def _start_heartbeat():
    import threading as _t, time as _time, os as _os, io as _io
    def _beat():
        while True:
            try:
                last = ''
                try:
                    with _io.open(LOG_PATH, 'r', encoding='utf-8') as f:
                        _lines = f.read().splitlines()
                        last = _lines[-1] if _lines else ''
                except Exception:
                    pass
                with _io.open(HEARTBEAT_PATH, 'w', encoding='utf-8') as f:
                    f.write('%s | pid=%d | alive\nlast: %s\n' % (
                        _time.strftime('%m-%d %H:%M:%S'), _os.getpid(), last[:150]))
            except Exception:
                pass
            _time.sleep(5.0)
    _t.Thread(target=_beat, daemon=True, name='gui_heartbeat').start()


def log(s):
    _file_log(s)  # 先落盘：即使后续 print 阻塞，磁盘日志也不受影响
    print(s)
    if text_log:
        try:
            _log_queue.put_nowait(str(s))
        except Exception:
            text_log.insert(tk.END, str(s) + NL)

# ============================================================
# 连接（只连一次，复用）
# ============================================================
def ensure_connected():
    global _connected
    try:
        status, msg = robot.ConnectedState()
        if status != ROBOTCOM_READY:
            if status >= 0:
                log('机器人未就绪，取消执行：' + str(msg))
                return False
            robot.Connect()
            # v14o：固定 1.5s 改为就绪探测（0.3s 轮询，最多 3s）：假断连恢复是每跳尾部
            # 停顿税的一部分；探测到就绪即返回，未就绪语义与旧版一致（返回 False）。
            for _ in range(10):
                time.sleep(0.3)
                status, msg = robot.ConnectedState()
                if status == ROBOTCOM_READY:
                    break
        _connected = status == ROBOTCOM_READY
        if not _connected:
            log('机器人连接未就绪：' + str(msg))
            return False
        RDK.setRunMode(RUNMODE_RUN_ROBOT)
        return True
    except Exception as exc:
        _connected = False
        log('连接失败：' + str(exc))
        return False


# ============================================================
# 解析坐标
# ============================================================
def parse_points():
    if not text_points:
        return []
    raw = text_points.get("1.0", tk.END)
    points = []
    for line in raw.strip().split(NL):
        line = line.strip()
        if not line or line.startswith("#"):
            continue
        try:
            vals = [float(v.strip()) for v in line.split(",")]
            if len(vals) >= 6:
                points.append(vals[:6])
        except ValueError:
            pass
    return points

# ============================================================
# 读取当前位置
# ============================================================
def read_current(entries=None):
    try:
        pose = robot.Pose()
        v = pose_to_fanuc(pose)
        log("")
        log("当前 TCP：X=%.3f Y=%.3f Z=%.3f Rx=%.3f Ry=%.3f Rz=%.3f" % tuple(v[:6]))
    except Exception as e:
        log("读取失败：%s" % e)

def fill_current(entries=None):
    try:
        pose = robot.Pose()
        v = pose_to_fanuc(pose)
        if entries:
            for e, val in zip(entries, v):
                e.delete(0, tk.END)
                e.insert(0, "%.3f" % val)
        log("当前 TCP 已填入")
    except Exception as e:
        log("读取失败：%s" % e)

# ============================================================
# IK 检测
# 注意：SolveIK 显式使用当前 Tool + Reference，和 MoveL/MoveJ 保持一致。
# ============================================================
def check_ik_single(entries=None):
    if not entries:
        return
    try:
        values = [float(e.get()) for e in entries]
    except ValueError:
        log("输入无效")
        return

    x, y, z, rx, ry, rz = values
    target = fanuc_to_pose(x, y, z, rx, ry, rz)
    log("")
    log("目标：X=%.3f Y=%.3f Z=%.3f Rx=%.3f Ry=%.3f Rz=%.3f" % (x, y, z, rx, ry, rz))

    try:
        tool_pose = robot.PoseTool()
        frame_pose = robot.PoseFrame()
        joints = robot.SolveIK(target, tool=tool_pose, reference=frame_pose)
        if joints is None:
            log("IK 不可达")
        else:
            q = joints.list()
            if len(q) < 6:
                log("IK 返回关节数量异常：%d，原始数据=%r" % (len(q), q))
                return
            log("IK 可达")
            log("  关节：J1=%.2f J2=%.2f J3=%.2f J4=%.2f J5=%.2f J6=%.2f" % tuple(q[:6]))
    except Exception as e:
        log("检测失败：%s" % e)

def check_all_ik():
    points = parse_points()
    if not points:
        log("没有有效点")
        return

    log("")
    log("========== 检测全部 %d 个点 ==========" % len(points))
    all_ok = True
    for i, p in enumerate(points):
        try:
            target = fanuc_to_pose(*p)
            joints = robot.SolveIK(target, tool=robot.PoseTool(), reference=robot.PoseFrame())
            if joints is None:
                log("  P%d: 不可达" % (i+1))
                all_ok = False
            else:
                q = joints.list()
                if len(q) < 6:
                    raise ValueError("IK 返回关节数量异常: %d, raw=%r" % (len(q), q))
                log("  P%d: 可达  J1=%.1f J2=%.1f J3=%.1f J4=%.1f J5=%.1f J6=%.1f" % (i+1, *q[:6]))
        except Exception as e:
            log("  P%d: 检测失败 %s" % (i+1, e))
            all_ok = False
    if all_ok:
        log("全部 %d 个点可达" % len(points))
    else:
        log("存在不可达点，执行前整段预检将拒绝不通过的方案")

# ============================================================
# 执行单点
# ============================================================
def execute_single(entries=None, mtype="MoveL"):
    try:
        if not entries:
            return
        values = [float(e.get()) for e in entries]
        _execute_checked_real([dict(type='TCP', values=values)], single_method=mtype)
    except (ValueError, TypeError) as exc:
        log('单点输入无效：' + str(exc))


# ============================================================
# 连续运动：选项卡3直接输入 TCP / 关节点，逐点检查后加入轨迹
# ============================================================
trajectory_records = []
record_text = None
traj_entries = None
traj_type = None
singular_var = None
j6_direction_var = None
spin_var = None


def _parse_six_from_entries(entries, label):
    if not entries or len(entries) != 6:
        log("%s输入框异常：需要 6 个值" % label)
        return None
    try:
        vals = [float(e.get().strip()) for e in entries]
    except (ValueError, AttributeError):
        log("%s输入无效：6 个值必须全部为数字" % label)
        return None
    if not all(math.isfinite(v) for v in vals):
        log("%s输入无效：不能包含 NaN 或无穷值" % label)
        return None
    return vals


def _check_tcp_reachable(vals):
    """检查单个 TCP 点 IK 是否可达，返回 (True, target, joints)。"""
    try:
        target = fanuc_to_pose(*vals)
        tool_pose = robot.PoseTool()
        frame_pose = robot.PoseFrame()
        joints = robot.SolveIK(target, tool=tool_pose, reference=frame_pose)

        if joints is None:
            log("TCP IK：不可达")
            return False, None, None

        q = joints.list()
        if len(q) < 6:
            log("TCP IK：返回关节数量异常：%r" % q)
            return False, None, None

        log("TCP IK：可达")
        log("  IK关节：J1=%.2f J2=%.2f J3=%.2f J4=%.2f J5=%.2f J6=%.2f" % tuple(q[:6]))
        return True, target, q[:6]
    except Exception as e:
        log("TCP IK 检查失败：%s: %s" % (type(e).__name__, e))
        return False, None, None


def _check_tcp_segment_continuous(prev_vals, curr_vals, segment_index, samples=20):
    """检查前一个 TCP 点到当前 TCP 点之间的整段插补路径 IK 连续可达性。

    暂不考虑障碍物，只对 TCP 位姿做线性插值，并对每个采样位姿执行 SolveIK。
    起点和终点也包含在采样检查中。
    """
    if prev_vals is None:
        return True

    log("开始检查 P%d -> P%d 的 TCP 连续 IK（%d 个采样点）" %
        (segment_index - 1, segment_index, samples + 1))

    tool_pose = robot.PoseTool()
    frame_pose = robot.PoseFrame()

    for k in range(samples + 1):
        t = float(k) / float(samples)
        vals = [prev_vals[i] + (curr_vals[i] - prev_vals[i]) * t for i in range(6)]
        try:
            pose = fanuc_to_pose(*vals)
            joints = robot.SolveIK(pose, tool=tool_pose, reference=frame_pose)
            if joints is None:
                log("  P%d -> P%d：第 %d/%d 个采样点 IK 不可达，t=%.3f" %
                    (segment_index - 1, segment_index, k + 1, samples + 1, t))
                log("  TCP：X=%.3f Y=%.3f Z=%.3f Rx=%.3f Ry=%.3f Rz=%.3f" % tuple(vals))
                return False
            q = joints.list()
            if len(q) < 6:
                log("  P%d -> P%d：第 %d 个采样点 IK 返回异常：%r" %
                    (segment_index - 1, segment_index, k + 1, q))
                return False
        except Exception as e:
            log("  P%d -> P%d：第 %d 个采样点 IK 检查失败：%s: %s" %
                (segment_index - 1, segment_index, k + 1, type(e).__name__, e))
            return False

    log("P%d -> P%d：连续 IK 检查通过" % (segment_index - 1, segment_index))
    return True


def _check_joint_reachable(q):
    """兼容旧代码：关节点不做可达性/限位检查，输入合法即可加入。"""
    return True


def refresh_record_list():
    if record_text is None:
        return

    record_text.delete("1.0", tk.END)

    for i, rec in enumerate(trajectory_records, 1):
        kind = rec["type"]
        vals = rec["values"]

        if kind == "TCP":
            if rec.get("spin360", False):
                mark = " [J6自转360° %s]" % ("+" if rec.get("j6_delta", 360) >= 0 else "-")
            elif rec.get("singular", False):
                mark = " [J6特异点 %s180°]" % ("+" if rec.get("j6_delta", 180) >= 0 else "-")
            else:
                mark = ""
            record_text.insert(
                tk.END,
                "P%-3d [TCP]%s   X=%9.3f Y=%9.3f Z=%9.3f Rx=%8.3f Ry=%8.3f Rz=%8.3f%s" %
                (i, mark, *vals, NL)
            )
        else:
            record_text.insert(
                tk.END,
                "P%-3d [JNT]   J1=%8.3f J2=%8.3f J3=%8.3f J4=%8.3f J5=%8.3f J6=%8.3f%s" %
                (i, *vals, NL)
            )


def add_and_check_trajectory_point():
    values = _parse_six_from_entries(traj_entries, traj_type.get())
    if values is None:
        return
    kind = traj_type.get()
    is_singular = kind == 'TCP' and bool(singular_var.get())
    spin = is_singular and bool(spin_var.get())
    sign = 1 if int(j6_direction_var.get()) >= 0 else -1
    rec = dict(type=kind, values=values, singular=is_singular, spin360=spin,
               j6_delta=sign * (360 if spin else 180))
    try:
        records = _validated_records(trajectory_records + [rec])
    except ValueError as exc:
        log('点未加入：' + str(exc))
        return
    trajectory_records[:] = records
    refresh_record_list()
    if spin:
        log('P%d [TCP-J6自转360°]：已加入；执行时 J1~J5 不变，J6 %+d°。' % (len(records), sign * 360))
    else:
        log('点已加入；完整避障预检将在执行前进行。关节圈数按输入保留。')



def _write_values_to_traj_entries(values, label):
    if not traj_entries or len(traj_entries) != 6:
        log("连续运动输入框异常：无法写入当前%s" % label)
        return False
    for e, val in zip(traj_entries, values[:6]):
        e.delete(0, tk.END)
        e.insert(0, "%.3f" % float(val))
    log("当前%s已写入选项卡3输入框" % label)
    return True


def read_current_tcp_to_traj():
    """读取当前 RoboDK TCP，并写入选项卡3的 TCP 输入框。"""
    try:
        pose = robot.Pose()
        vals = pose_to_fanuc(pose)
        log("========== 读取当前 TCP -> 选项卡3 ==========")
        log("X=%+.3f Y=%+.3f Z=%+.3f Rx=%+.3f Ry=%+.3f Rz=%+.3f" % tuple(vals))
        if traj_type.get() != "TCP":
            traj_type.set("TCP")
            _update_traj_labels_and_defaults()
        return _write_values_to_traj_entries(vals, "TCP")
    except Exception as e:
        log("读取当前 TCP 失败：%s: %s" % (type(e).__name__, e))
        return False


def read_current_joints_to_traj():
    """读取 RoboDK Robot Item 当前关节，并写入选项卡3的关节输入框。"""
    q = read_current_joints(None)
    if q is None or len(q) < 6:
        return False
    log("========== 读取当前关节 -> 选项卡3 ==========")
    if traj_type.get() != "JOINT":
        traj_type.set("JOINT")
        _update_traj_labels_and_defaults()
    return _write_values_to_traj_entries(q, "关节")


def clear_trajectory_input():
    if not traj_entries:
        return

    for e in traj_entries:
        e.delete(0, tk.END)

    if traj_type.get() == "TCP":
        defaults = ["0.000", "-241.500", "1047.000", "-90.000", "0.000", "180.000"]
    else:
        defaults = ["0.000"] * 6

    for e, val in zip(traj_entries, defaults):
        e.insert(0, val)




def import_trajectory():
    filepath = filedialog.askopenfilename(title='导入轨迹', defaultextension='.json', filetypes=[('JSON轨迹','*.json'),('所有文件','*.*')])
    if not filepath:
        return
    try:
        with open(filepath, encoding='utf-8') as f:
            records = _validated_records(json.load(f))
        trajectory_records[:] = records
        refresh_record_list()
        log(f'已导入{len(records)}点：{filepath}。执行前将从实机当前关节重新预检。')
    except Exception as exc:
        log('轨迹导入失败：' + str(exc))


def delete_last_record():
    if trajectory_records:
        rec = trajectory_records.pop()
        refresh_record_list()
        log("已删除最后一点：P%d [%s]" %
            (len(trajectory_records) + 1, rec["type"]))
    else:
        log("当前没有可删除的连续运动点")


def clear_records():
    trajectory_records.clear()
    refresh_record_list()
    log("连续运动点列表已清空")


def execute_recorded_trajectory():
    log('【点击】执行整段连续运动：当前列表 %d 点（转后台线程执行，窗口保持响应）' % len(trajectory_records))
    import threading
    def _worker():
        try:
            _execute_checked_real(list(trajectory_records))
        except Exception as exc:
            log('【线程异常】%s: %s' % (type(exc).__name__, exc))
    threading.Thread(target=_worker, daemon=True, name='real_exec').start()



# 保留旧函数名，避免其他代码调用失效。
def execute_trajectory():
    execute_recorded_trajectory()


# ============================================================
# 实机关节运动
# ============================================================
def _joint_values_from_entries(entries):
    """从 GUI 读取 J1~J6 目标角度。单位：deg。"""
    if not entries or len(entries) != 6:
        log("目标关节输入框异常：需要 J1~J6 共 6 个")
        return None
    try:
        q = [float(e.get().strip()) for e in entries]
    except (ValueError, AttributeError):
        log("目标关节输入无效：J1~J6 必须全部填写数字")
        return None
    if not all(math.isfinite(v) for v in q):
        log("目标关节输入无效：不能包含 NaN 或无穷值")
        return None
    return q


def read_current_joints(entries=None):
    """读取 RoboDK Robot Item 当前关节值，并可直接填入 J1~J6 输入框。
    注意：这里读取的是 RoboDK 当前 Robot Item 的关节状态，不调用 CR5 控制器 GetAngle。
    """
    try:
        joints = robot.SimulatorJoints()
        q = list(joints) if hasattr(joints, "__iter__") else [joints]
        if len(q) < 6:
            log("读取当前关节失败：SimulatorJoints 返回 %r" % (q,))
            log("请确认 RoboDK 窗口中的机器人已经连接并显示实时关节角度。")
            return None

        q = q[:6]
        log("")
        log("========== RoboDK 当前关节 ==========")
        log("J1=%+.3f°  J2=%+.3f°  J3=%+.3f°" % tuple(q[:3]))
        log("J4=%+.3f°  J5=%+.3f°  J6=%+.3f°" % tuple(q[3:]))

        if entries and len(entries) == 6:
            for e, val in zip(entries, q):
                e.delete(0, tk.END)
                e.insert(0, "%.3f" % val)
            log("当前关节已填入 J1~J6 输入框")

        return q
    except Exception as e:
        log("读取 RoboDK 当前关节失败：%s: %s" % (type(e).__name__, e))
        return None


def fill_current_joints(entries=None):
    """当前 RoboDK 关节 -> 目标关节输入框。"""
    return read_current_joints(entries)


def execute_joint_target(entries=None):
    q = _joint_values_from_entries(entries)
    if q is not None:
        _execute_checked_real([dict(type='JOINT', values=q)])



def clear_joint_target(entries=None):
    if not entries:
        return
    for e in entries:
        e.delete(0, tk.END)
        e.insert(0, "0.000")
    log("目标关节输入已清零")

# ============================================================
# GUI
# ============================================================

# 与TCP仿真一致的预检核心；仅在仿真模式调用。
fanuc_values_to_pose = fanuc_to_pose
pose_to_fanuc_values = pose_to_fanuc
MOVEJ_FALLBACK_MAX_DEVIATION_MM = 50.0
# 预检缓存（与TCP仿真副本同款）：生命周期=单次预检规划，_enable_obstacle_checks 每次进入预检时清空。

_plan_cache = {}
_preferred_seed = None  # Ordering hint only; never reuse a collision certificate.


def _lazy_valid_seeds(seeds, start):
    """Keep the existing valid-seed order, testing only seeds actually needed.

    If none is reachable, preserve the old fallback to the unfiltered list.
    """
    found = False
    for seed in seeds:
        if seed is None or _movej_test_cached(start, seed, 1) == 0:
            found = True
            yield seed
    if not found:
        yield from seeds

def _cache_key_joints(q):
    return tuple(round(float(v), 3) for v in q[:6])

def _cache_key_pose(pose):
    return tuple(tuple(round(float(v), 6) for v in row) for row in pose.rows)

def _movej_test_cached(start, end, minstep_deg):
    """robot.MoveJ_Test 的缓存包装，返回值与直接调用完全一致。
    成功时与原调用一样把仿真关节停在终点；失败路径的规划器只依赖局部
    关节变量（不读取此时的模型关节状态），无需复现失败的副作用。"""
    key = ('movej_test', _cache_key_joints(start), _cache_key_joints(end),
           round(float(minstep_deg), 6))
    if key not in _plan_cache:
        _plan_cache[key] = robot.MoveJ_Test(start, end, minstep_deg=minstep_deg)
    elif _plan_cache[key] == 0:
        robot.setJoints(list(end[:6]))
    return _plan_cache[key]

def _tcp_target_to_flange(target):
    """输入是参考系中的TCP；IK需要机器人基座系中的法兰位姿。"""
    return robot.PoseFrame() * target * invH(robot.PoseTool())

def _flange_target_description(target):
    flange = _tcp_target_to_flange(target)
    return ('换算后的法兰中心（基座系）XYZ=' +
            str(tuple(round(v, 3) for v in flange.Pos())) +
            ' mm，法兰Z轴方向=' + str(tuple(round(v, 6) for v in flange.VZ())))


def _validated_records(data):
    if not isinstance(data, list) or not data:
        raise ValueError('轨迹必须是非空点列表。')
    result = []
    for i, rec in enumerate(data, 1):
        kind = str(rec.get('type', '')).upper()
        if kind == 'JNT':
            kind = 'JOINT'
        values = [float(v) for v in rec.get('values', [])]
        if kind not in ('TCP', 'JOINT') or len(values) != 6 or not all(math.isfinite(v) for v in values):
            raise ValueError(f'P{i}：类型或六维数值无效。')
        special = bool(rec.get('singular', False)) and kind == 'TCP'
        spin = special and bool(rec.get('spin360', False))
        raw_delta = int(rec.get('j6_delta', 360 if spin else 180)) if special else 0
        if special and (not result or result[-1]['type'] != 'TCP' or result[-1]['singular']):
            raise ValueError(f'P{i}：特异点前序或转向无效。')
        if special:
            if spin:
                if raw_delta not in (-360, 360):
                    raise ValueError(f'P{i}：J6自转方向必须为+360或-360。')
                if max(abs(a - b) for a, b in zip(values, result[-1]['values'])) > 1e-3:
                    raise ValueError(f'P{i}：J6自转360°特异点的六维数值必须与前一个TCP点完全相同。')
            elif raw_delta not in (-180, 180):
                raise ValueError(f'P{i}：J6方向必须为+180或-180。')
        delta = (360 if spin else 180) * (1 if raw_delta >= 0 else -1) if special else 0
        result.append(dict(type=kind, values=values, singular=special, spin360=spin, j6_delta=delta))
    return result


def _controller_feedback():
    # Dobot CR V3: 1440-byte real-time feedback; no command is sent on this socket.
    import socket
    import struct
    host, port, *_ = robot.ConnectionParams()
    if int(port) != 29999:
        raise RuntimeError('当前连接不是已验证的Dobot CR反馈协议。')
    previous = None
    with socket.create_connection((host, 30004), timeout=3.0) as connection:
        deadline = time.monotonic() + 3.0
        for _ in range(2):
            packet = bytearray()
            while len(packet) < 1440:
                remaining = deadline - time.monotonic()
                if remaining <= 0:
                    raise RuntimeError('实机反馈读取超时。')
                connection.settimeout(remaining)
                part = connection.recv(1440 - len(packet))
                if not part:
                    raise RuntimeError('实机反馈连接已关闭。')
                packet.extend(part)
            length = struct.unpack_from('<Q', packet, 0)[0]
            marker = struct.unpack_from('<Q', packet, 48)[0]
            stamp = struct.unpack_from('<Q', packet, 32)[0]
            if length != 1440 or marker != 0x123456789ABCDEF:
                raise RuntimeError('实机反馈帧格式不匹配。')
            if previous is not None and stamp <= previous:
                raise RuntimeError('实机反馈时间戳未更新。')
            previous = stamp
        q = list(struct.unpack_from('<6d', packet, 192))   # ★真实关节角（v10定位，示教器交叉证实）；旧版误读432="连接基准+指令累加"的假值
        velocity = list(struct.unpack_from('<6d', packet, 480))
        mode = struct.unpack_from('<Q', packet, 24)[0]
        if not all(math.isfinite(v) for v in q + velocity):
            raise RuntimeError('实机反馈包含无效关节数值。')
        return q, velocity, mode


def _live_joints():
    if RDK.RunMode() != RUNMODE_RUN_ROBOT:
        raise RuntimeError('当前不是实机执行模式。')
    status, msg = robot.ConnectedState()
    if status != ROBOTCOM_READY:
        raise RuntimeError('机器人未就绪或已断连：' + str(msg))
    q, velocity, mode = _controller_feedback()
    # 阈值由 0.1 放宽到 1.0：实测静止时 J4/J3 的速度估计噪声可达 0.31°/s
    # （六轴角度 8 次采样完全相同），0.1 会把"其实已静止"误判为运动中而中止任务。
    if mode != 5 or max(abs(v) for v in velocity) > 1.0:
        raise RuntimeError('实机未处于使能静止状态，模式=%s。' % mode)
    return q


def _require_joints(expected, _tries=3, _allow_fix=False):
    """校验关节与预检一致（容差 0.5°）；失败时【主动发一条 MoveJ 校正】，仍不行才抛错。

    ★★★ v15.10（2026-11-03）：根治"走到 P8 后不动"。
    根因（读码确认）：`_settle_core` 的断连分支写的是
        `_wait_arrival_then_static(expect_target)`
      · 直发段传了 expect_target ⇒ 会等到目标 ✓
      · **MoveJ 段传的是 None** ⇒ 退化为「只等静止」✗
      ⇒ 指令被断连打断、手臂停在中途 ⇒ 只要「静止」就算完成 ✗
      ⇒ 下一段开头的 _require_joints 发现差 9.77° ⇒ 抛错 ⇒ 停 ✗
    （历史证据：10-13 12:12 / 15:49 / 15:55 三次同样失败，当时 P8 走的是纯 MoveJ，与直发无关 ✗）

    修法：不再是"发现不一致就停"，而是【发一条 MoveJ 到认证关节】把手臂拉回去，再校验。
      · 目标就是预检认证过的关节构型 ⇒ 确定可达 ⇒ 重发安全 ✓
      · 只补一次（_allow_fix=False 时不再递归）⇒ 不会无限循环 ✓
      · 拉回后仍不一致 ⇒ 才抛错 ✓（护栏不放松）
    """
    last = None
    actual = None
    for k in range(_tries):
        actual = _live_joints()
        last = max(abs(a - b) for a, b in zip(actual, expected))
        if last <= 0.5:
            return
        if k < _tries - 1:
            log('关节偏差 %.2f° > 0.5°（第 %d/%d 次）⇒ 等 0.5s 重读（可能仍在微动）'
                % (last, k + 1, _tries))
            time.sleep(0.5)
    if _allow_fix:
        log('关节偏差 %.2f°（目标%s，实测%s）⇒ 主动发 MoveJ 校正到认证关节（v15.10）'
            % (last, ['%.2f' % v for v in expected], ['%.2f' % v for v in (actual or [])]))
        try:
            robot.MoveJ(list(expected))
            time.sleep(1.0)
            _require_joints(expected, _tries=3, _allow_fix=False)
            log('✓ 校正 MoveJ 生效：关节已回到认证构型')
            return
        except Exception as _fix_exc:  # noqa: BLE001
            log('⚠️ 校正 MoveJ 未生效：%s: %s' % (type(_fix_exc).__name__, _fix_exc))
    raise RuntimeError('关节反馈与预检状态不一致（偏差 %.2f°，目标%s，实测%s），停止后续命令。'
                       % (last, ['%.2f' % v for v in expected], ['%.2f' % v for v in (actual or [])]))


def _retreat_orientation_records(records):
    """加工点变姿态前退到 y=-750，变姿态后返回 y=-775。"""
    result = []
    previous = None
    for index, record in enumerate(records, 1):
        current = dict(record, values=record['values'][:])
        current['label'] = f'P{index}'
        if previous and previous['type'] == current['type'] == 'TCP':
            old, new = previous['values'], current['values']
            changed = pose_angle(invH(fanuc_values_to_pose(*old)) * fanuc_values_to_pose(*new)) > math.radians(.01)
            old_work, new_work = abs(old[1] + 775) < .001, abs(new[1] + 775) < .001
            if changed and (old_work or new_work):
                anchor = old if old_work else new
                retreat = dict(type='TCP', values=[anchor[0], -750., anchor[2]] + old[3:], singular=False,
                               label=f'P{index}前退让', require_linear=old_work)
                result.append(retreat)
                turn = dict(current, values=retreat['values'][:3] + new[3:], label=f'P{index}退让位换向')
                result.append(turn)
                current['singular'] = False
                current['require_linear'] = new_work
        result.append(current)
        previous = record
    return result


def _prepare_real_plan(records, start, deviation, single_method=None):
    RDK.setRunMode(RUNMODE_SIMULATE)
    try:
        RDK.Command('Trace', 'Off')
        robot.setJoints(start)
        if single_method is None:
            return _plan_continuous_trajectory(records, deviation, log)
        _enable_obstacle_checks()
        if robot.MoveJ_Test(start, start, minstep_deg=1) != 0:
            raise ValueError('起始姿态碰撞：' + _collision_details())
        values = records[0]['values']
        method, fallback = single_method, False
        if method not in ('MoveJ','MoveL'):
            raise ValueError('未知单点运动类型。')
        end = None
        waypoints = []
        if method == 'MoveL':
            end, _ = _linear_path_endpoint(start, fanuc_to_pose(*values))
            if end is not None:
                # v13：单点 MoveL 同样不信任驱动 MOVL（纯J6自转也一样，关节插值=同一路径），
                # 改细分途经点+MoveJ 执行
                waypoints = _linear_waypoints(start, fanuc_to_pose(*values))
                if waypoints:
                    log('单点 MoveL 改细分执行：%d 个途经点（步长≤%.0fmm）。' % (len(waypoints), LINEAR_SUBSTEP_MM))
                    log('单点 MoveL 途经跳（共%d跳）：%s' % (len(waypoints), [[float('%.2f' % v) for v in w] for w in waypoints]))
        if end is None:
            end = _obstacle_joint_target(start, values, deviation if method=='MoveL' else None)
            fallback, method = method=='MoveL', 'MoveJ'
        plan = [dict(method=method,joints=end,special=False,fallback=fallback,rewinds=[],j6_delta=None,waypoints=waypoints)]
        _verify_obstacle_plan(start, plan)
        return plan
    finally:
        robot.setJoints(start)
        RDK.Render(True)
        RDK.setRunMode(RUNMODE_RUN_ROBOT)  # 旧版 L615 有此行：预检后必须切回实机模式，否则 _live_joints 直接拒执行


def _wait_controller_static(max_wait_s=20.0, vel_threshold=0.5, samples=5, interval=0.3):
    """轮询30004反馈直到六轴静止（连续samples次速度<阈值），返回(关节, 是否静止)。

    v14o：断连分支以 samples=3/interval=0.2 调用（短跳≈1s，5×0.3s 静止确认占每跳
    尾部 ~1.5s，是停顿税大头）；默认 5×0.3s 供正常路径；20s 静止上限（真断连护栏）不动。"""
    t0 = time.time()
    quiet = 0
    last = None
    while time.time() - t0 < max_wait_s:
        actual, velocity, _mode = _controller_feedback()
        last = actual
        if max(abs(v) for v in velocity) < vel_threshold:
            quiet += 1
            if quiet >= samples:
                return last, True
        else:
            quiet = 0
        time.sleep(interval)
    return last, False


class ControllerMotionFault(RuntimeError):
    """A controller state that must never trigger a motion resend."""
    pass


def _wait_arrival_then_static(target_joints, max_wait_s=20.0):
    """v14u：目标锚定的到位等待——直发后不再猜「起步了没」，只等「到没到」。

    背景（v14t 10:38 P9 实测）：直发指令起步延迟可 >6s，让位 6s 耗尽判「未执行」
    停止后，指令仍被控制器自行执行到精确目标（善后实测 J2 +10°/J3 +20°，余轴不动，
    宏未重发）——「起点静止」与「完成静止」在反馈上不可区分，位置对目标才是唯一
    可靠锚点（速度判据出局：三场停时 J4 0.06~0.42°/s 均为低于阈值的保持抖动）。
    本函数：距目标关节 ≤MOVL_ARRIVE_TOL_DEG 且速度<0.5°/s → 到位完成（此时已在
    目标，无需再做常规静止确认）；每 5s 一行进度日志（顺带实测真实延迟）；
    上限 MOVL_ARRIVE_WAIT_S 超时报「疑似未执行」停待判读；不重发铁律不变。
    target_joints=None → 退化为 _wait_controller_static()，行为与原先完全一致。"""
    if target_joints is not None:
        t0 = time.time()
        t_note = t0
        while True:
            fb = _controller_feedback()
            if fb[2] not in (5, 7, 8):
                raise ControllerMotionFault(
                    '控制器反馈模式=%s，停止等待且不补发；目标关节=%s，实际关节=%s。请检查示教器报警。'
                    % (fb[2], target_joints, fb[0]))
            err = max(abs(a - b) for a, b in zip(fb[0], target_joints))
            if err <= MOVL_ARRIVE_TOL_DEG and max(abs(v) for v in fb[1]) < 0.5:
                log('MovL 直发到位确认：距目标关节%.2f°（%.1fs），验收继续。'
                    % (err, time.time() - t0))
                return fb[0], True
            if time.time() - t0 >= MOVL_ARRIVE_WAIT_S:
                raise RuntimeError(
                    'MovL 直发%.0fs仍未到位（距目标关节%.2f°），疑似未执行，停止待判读。'
                    % (MOVL_ARRIVE_WAIT_S, err))
            if time.time() - t_note >= 5.0:
                log('MovL 直发等待到位：%.0fs，距目标关节%.2f°，续等（不重发，上限%.0fs）。'
                    % (time.time() - t0, err, MOVL_ARRIVE_WAIT_S))
                t_note = time.time()
            time.sleep(0.5)
    return _wait_controller_static(max_wait_s=max_wait_s)


MOVE_OFFSET_TOL = 0.5   # 闭环补偿后的到位容差（°）


TCP_TOOL_NAME = 'CR5_TCP_130mm'
FLANGE_TOOL_NAME = '_CR5_FLANGE_DIRECT_TEMP'
_tool_window_depth = 0


def _same_tool_pose(a, b):
    return max(abs(a[r, c] - b[r, c]) for r in range(4) for c in range(4)) < 1e-7


def _named_tool(name, pose):
    matches = [it for it in robot.Childs()
               if it.Type() == ITEM_TYPE_TOOL and it.Name() == name]
    if len(matches) > 1:
        raise RuntimeError('重复 TCP 工具条目：' + name)
    if matches:
        tool = matches[0]
        if not _same_tool_pose(tool.PoseTool(), pose):
            raise RuntimeError('TCP 工具定义不符，停止待核对：' + name)
        return tool
    return robot.AddTool(pose, name)


def _restore_tool(pose, linked_tool=None):
    """Restore the original item link when possible, and never swallow failure."""
    for attempt in range(2):
        try:
            robot.setPoseTool(linked_tool if linked_tool is not None and linked_tool.Valid() else pose)
            if not _same_tool_pose(robot.PoseTool(), pose):
                raise RuntimeError('PoseTool 恢复后读回不一致')
            return
        except Exception as exc:
            if attempt == 1:
                raise RuntimeError('工具恢复失败，禁止继续运动：' + str(exc)) from exc


def _single_move_settle(method, target, require_joints=True, expect_target=None, flange_space=False, _retry=0):
    """发指令并确认到位——v14w39 窗口版入口：flange_space 时单位变换+藏把手覆盖
    【整个 settle 生命周期】（发送+断连恢复+到位等待）。旧版只包 RPC 一次调用：假断连
    抛出时窗口即关、把手提前回来，RoboDK 本地退化动画在弧 66% 被碰撞检测掐停→模型冻在
    撞点、红显常驻→收口 MoveJ 被拦死（10-22 四次实录含 v14w38）。"""
    global _tool_window_depth
    if not flange_space or _tool_window_depth:
        # A controlled retry already runs inside the outer tool window.
        # Only the outer owner may restore the original TCP.
        return _settle_core(method, target, require_joints, expect_target, flange_space, _retry)
    _ensure_canonical_tool()
    _win_tp = robot.PoseTool()
    _win_link = robot.getLink(ITEM_TYPE_TOOL)
    _win_handle = RDK.Item('门把手_bs1')
    _win_visible = _win_handle.Visible() if _win_handle.Valid() else None
    _flange_tool = _named_tool(FLANGE_TOOL_NAME, eye(4))
    _tool_window_depth += 1
    try:
        robot.setPoseTool(_flange_tool)
        if not _same_tool_pose(robot.PoseTool(), eye(4)):
            raise RuntimeError('法兰工具切换失败，未发送运动指令')
        if _win_visible is not None:
            _win_handle.setVisible(False)
        result = _settle_core(method, target, require_joints, expect_target, True, _retry)
        # Synchronize measured joints before restoring the tool and visible mesh.
        actual, is_static = _wait_controller_static()
        if not is_static:
            raise RuntimeError('法兰直发后未确认静止，停止后续命令。')
        robot.setJoints(actual)
        return result
    finally:
        try:
            _restore_tool(_win_tp, _win_link)
        finally:
            _tool_window_depth -= 1
            if _win_visible is not None:
                _win_handle.setVisible(_win_visible)


def _settle_core(method, target, require_joints, expect_target, flange_space=False, _retry=0):
    """发一条运动指令并确认到位（v10：反馈字段已校正）。

    v14r：require_joints=False 仅供 MovL 直发调用点使用——断连分支的关节级 0.5°
    校验让位给外层法兰级粗验收（≤8mm/≤1°）+MoveJ 微纠偏收口（v14q 09:57 实机
    教训：MovL 直发必触发假断连，0.95° 固有残差在断连分支内即被拦停，外层验收
    根本没执行到）。其余护栏不变：20s 静止上限、重连失败仍停。

    v14u：断连分支改目标锚定到位等待 _wait_arrival_then_static——上限 60s 每 5s
    进度日志；超时报「疑似未执行」停。不重发铁律不变。

    v14w37：直发=【法兰位姿传递 + flange_space 单位变换窗口】双件套——
    ①传位姿（调用方 invH(PoseFrame)*SolveFK(净化关节) 自算）：MoveL 的动画按位姿空间
    直线走=认证路径，根治旧 MoveL(关节) 的关节弧动画扫进圆柱假碰撞冻死（10-22 两次实录）；
    ②发送 RPC 窗口内 PoseTool 置单位变换：MoveL(位姿) 的可达校验/语义都按 TCP 空间做，
    不切工具则法兰位姿被当 TCP 反推（P8 反推法兰 z=744 爆臂展 ⇒ TargetReachError，
    10-22 11:18 实录）；单位变换下校验空间=法兰空间，数字逐位=金标准（实证 0 偏差）。
    动画窗口内直线途经点 12/12 无碰撞（单位变换工具下实测）。
    v14w38：窗口内追加隐藏把手——驱动断连瞬间 RoboDK 本地退化关节动画（会撞圆柱的
    那条弧）是三次冻结的真凶；藏把手=对假路径的检测放行（实测弧中点/冻结姿态
    显隐 True/False 翻转），真直线 1mm 检查本来就 0 碰撞。

    v14w20：受控补发（一次性）——驱动连接恰死在发送时刻时 SendJointMovJ 会静默
    丢弃不发送（反汇编：CONNECTED=False 直接 return False；2026-10-15 09:51 P25
    实发：断连后臂停在发送前位置、误差127.8°）。补发条件（全部满足才补，且全程
    至多一次）：①失败 ②30004 独立反馈证明【零位移】（仍在发送前关节 ≤0.5°）
    ③ensure_connected() 重连成功。指令已上线/延迟执行/落点异常的场景均不满足
    ②（有位移）不会触发——保留原「不重发」语义。历史上"晚执行"案例（v14t）
    后经控制器日志证实为面板拖动误判，非队列延迟。

    历史结论：驱动一直正确执行绝对关节目标；真实关节角在偏移192。"""
    try:
        _start_q = None
        try:
            _start_q = _controller_feedback()[0]
        except Exception:
            _start_q = None
        getattr(robot, method)(target)   # v14w39：flange 窗口已上移至 _single_move_settle 包装层
    except StoppedError as exc:
        if str(exc).strip() != 'Robot not connected':
            raise
        # v14o 静默重连：假断连是本环境常态（每条 MoveJ 指令结束后都可能误报）；30004
        # 反馈通道独立于驱动连接，静止确认与重连并行进行，压缩跳间停顿税。
        # 护栏不变：未自然收尾（20s 上限）仍停、落点仍 0.5° 校验、重连失败仍停。
        log('驱动报断连——等待收尾与后台重连并行进行…')
        import threading as _st
        reconnected = []
        def _bg_reconnect():
            for _r in range(3):
                if ensure_connected():
                    reconnected.append(True)
                    return
                time.sleep(1.0)
        _rt = _st.Thread(target=_bg_reconnect, daemon=True, name='silent_reconnect')
        _rt.start()
        # v14u：到位等待下沉在断连分支（MovL 直发永远走本分支——v14s 教训）——
        # 目标锚定：距目标≤2°且静止=完成，不猜起步。非 MovL 直发退化为常规静止确认。
        try:
            actual, is_static = _wait_arrival_then_static(expect_target)
        except RuntimeError as _arr_exc:
            if isinstance(_arr_exc, ControllerMotionFault):
                raise
            # v14w20：直发「疑似未执行」——零位移+重连成功 ⇒ 补发一次（指令未上线实证）
            if (_retry < 1 and _start_q is not None
                    and max(abs(a - b) for a, b in zip(_controller_feedback()[0], _start_q)) <= MOVE_OFFSET_TOL
                    and ensure_connected()):
                log('直发疑似未执行且零位移（仍在起点）——判定指令未上线，补发一次（v14w20）。')
                return _single_move_settle(method, target, require_joints, expect_target,
                                           flange_space, _retry=_retry + 1)
            raise
        if not is_static:
            raise RuntimeError('驱动报断连后等待%.0fs仍未静止，停止。' % 20.0) from exc
        if require_joints:
            err = max(abs(a - b) for a, b in zip(actual, target))
            if err > MOVE_OFFSET_TOL:
                # v14w20：MoveJ 类「断连收尾后未到位」——零位移+重连成功 ⇒ 补发一次
                if (_retry < 1 and _start_q is not None
                        and max(abs(a - b) for a, b in zip(actual, _start_q)) <= MOVE_OFFSET_TOL
                        and ensure_connected()):
                    log('断连后零位移（仍在起点）——判定指令未上线，补发一次（v14w20）。')
                    return _single_move_settle(method, target, require_joints, expect_target,
                                               flange_space, _retry=_retry + 1)
                raise RuntimeError('断连收尾后未到位：目标%s，实测%s（误差%.2f°），停止待判读。'
                                   % (['%.2f' % v for v in target], ['%.2f' % v for v in actual], err)) from exc
        _rt.join(timeout=4.0)
        if not reconnected:
            raise RuntimeError('已到位但驱动重连失败，停止后续指令。') from exc
        log('驱动断连但运动已自然完成到位；已重连驱动，继续。')
        return
    actual, is_static = _wait_controller_static()
    if not is_static:
        raise RuntimeError('指令返回后等待静止超时（20s），停止。')
    if require_joints:
        err = max(abs(a - b) for a, b in zip(actual, target))
        if err > MOVE_OFFSET_TOL:
            raise RuntimeError('落点偏差%.2f°：目标%s，实测%s，停止待判读。'
                               % (err, ['%.2f' % v for v in target], ['%.2f' % v for v in actual]))
    return


MOVE_OFFSET_TOL = 0.5   # 到位容差（°）：反馈字段校正后，超过即停止待判读


# v13（方案B）：驱动 MOVL 执行层已判死（3 次实机断连指纹 + .pyc 反汇编直连无收尾），
# 所有 MoveL 执行全部替换为「细分途经点 + MoveJ」。作业面短段（≤ TRANSIT_DIRECT_MAX_MM）
# 用 MoveL 指令的 1mm 逆解采样出 ≤ LINEAR_SUBSTEP_MM 的途经关节序列，MoveJ 逐跳执行；
# 过渡段长段优先 MoveJ 直达（须过 TCP 偏离≤max_deviation 且整弧 MoveJ_Test 碰撞检查），
# 不满足才退回细分。预检层 MoveL_Test@1mm 保留：仍是「这一段能不能走直线」的权威筛选器。
TRANSIT_DIRECT_MAX_MM = 300.0   # 超过此段长的 TCP 段视为自由空间过渡段，尝试 MoveJ 直达
LINEAR_SUBSTEP_MM = 20.0        # 作业面细分步长：v14m(40mm) 实机碰撞实证弦误差可吃掉真裕度（轴线距199.9-半径180≈19.9mm），回 20mm 安全基准（v14k 两度全通过）；途经点弦误差 <0.5mm

MOVL_DIRECT_MAX_MM = 250.0   # v14w35（10-22）：150→210——150 是 v14p 照当时谱系（最长≈120mm）取的设计余量，非事故判死值；210 覆盖 200mm 工艺段一指令（y=-719 线翻转点→x=-100），留 FP 边界余量。路径背书不变（认证直线+整段复核）；更长直线段仍走细分
# ★★★ v14w（2026-10-13 16:08）：【禁直发名单清空 = 恢复 P9 直发】+ 发送位姿数字净化。
#   v14v4 按点号拦 P9 是在 -30001 真凶查明前的临时措施（且拦下分支会落空——随名单清空，
#   该落空分支变为不可达死码，留档不删）。真凶 = 控制器 MovL 参数校验拒收【参数形态】
#   （-0.000000 / +90.000000 / -0.000000，见 LOG_VERSION 处实录），不是几何、不是段长：
#   同目标 15:55:51 单步直发实证 return 0、1.1s 到位。净化失败 ⇒ 本段自动改走细分（安全回落）。
# 想再拦某点：改回 (9,) 即可（注意拦下分支的落空缺陷仍在，见 P2P_LESSONS.md）。
# ★★★ 2026-11-03：改回 (9,) —— 针对【新根因】"movL not set tool or user"（不是 -30001）
#   实录（控制器日志 11-03 10:33:24 / 10:33:30）：
#     [MovL#859] Motion args is legal!            ← 参数合法（所以不是 -30001）
#     [MovL#878] movL not set tool or user!!!     ← ★ 工具/用户坐标系没设置
#     [CallProcess#275] ret = 73/76 ... return = 0,{}  ← 被接受，但按【默认 tool/user】执行
#   ⇒ RoboDK 的 DobotCR 驱动下发 MovL(x,y,z,rx,ry,rz) 时【不带 tool/user】✗
#     ⇒ 控制器用开机默认值 ⇒ 与脚本"法兰补偿（PoseTool=eye）"的语义不一致 ⇒ 落点偏离（P9 差 11.80°）✗
#   ⇒ 保底：P9 不做直发，直接走【细分途经点路径】（今天 P5 就是这样走完的：13 途经点 ✓）
#   ⇒ 根治手段见下方 MOVL_SEND_TOOL_USER（实验性，默认关）
# ★★★ v15.9（2026-11-03）：P8 也加入禁直发 —— 直发的"选解自由"问题对 P8 同样致命。
#   实录（v15.8, 11:56:09~14）：
#     P8 直发 → 等静止 ✓ → 法兰验收通过（5.71mm/0.32° ✓）→ 收口 MoveJ
#     ⇒ 控制器最后停在【另一组 IK 解】：
#        目标 [68.33, 41.30, 10.92, 37.78, -90, 158.33]
#        实测 [78.10, 36.86, 19.48, 33.66, -90, 168.10]
#        差   +9.77, -4.44, +8.56, -4.12,  0,  +9.77
#     ⇒ J1 与 J6 同步 +9.77° ⇒ 【基座-腕部互相补偿】的同一法兰位姿、另一组解 ✗
#   ⇒ 根因：MovL 只给位姿 ⇒ 控制器自行选 IK 分支 ⇒ 关节构型不可控 ✗
#     （v15.5~v15.8 的等待/重试/安全网都改变不了这一点 ✗）
#   ⇒ 细分路径是【逐关节】走的 ⇒ 不存在选解问题 ⇒ 关节精确 ✓（代价：8 跳 ≈24 秒）
MOVL_DIRECT_BLOCK_POINTS = (9, 11)

# ★ 实验性开关（v15.3 已打开做验证）：直发前先给【控制器】发 Tool(0)/User(0)，
#   让 MovL 明确用 基座系+零工具(法兰)。背景：[MovL#878] movL not set tool or user!!!
#   ⇒ 控制器没收到 tool/user 就按默认执行 ⇒ 与"法兰补偿（PoseTool=eye）"语义不一致 ⇒ P9 落点偏 11.80°
#   验证目标：打开后控制器日志里 `movL not set tool or user` 是否消失。
#     消失 ⇒ 直发侧真能用 ⇒ "断断续续"（13 跳 × 3 秒）可根治 ✓
#     仍出现 ⇒ RoboDK DobotCR 驱动不透传 Tool()/User() ⇒ 此路不通，只能接受 3 秒/跳 ✗
#   安全性：发送失败只记日志、不阻断主流程；直发落点仍受法兰级粗验收（≤8mm/≤1°）护栏 ✓
MOVL_SEND_TOOL_USER = False  # RunCodeCustom is a project call, not raw dashboard transmission.
MOVL_FLANGE_TOL_MM = 8.0     # v14q 直发 MovL 法兰位置粗验收容差：控制器 MovL 固有落点残差实测 4.61mm（v14p 首航）/5.5mm（v14l）双样本，取实测+裕量；超此值=落点异常真停
MOVL_FLANGE_TOL_DEG = 1.0    # v14q 直发 MovL 法兰姿态粗验收容差（实测 0.616°+裕量）；通过后 MoveJ 微纠偏收口到关节级 0.5° 内
MOVL_ARRIVE_WAIT_S = 60.0    # v14u MovL 直发到位等待上限：目标锚定（距目标≤2°且静止即完成），不猜起步——v14t 10:38 实测 P9 起步延迟>6s、指令事后自行执行完；60s 为 10 倍裕量，每5s进度日志实测真实延迟，超时按未执行停待判读
MOVL_ARRIVE_TOL_DEG = 5.0    # v14u 到位判定关节距离阈（°）；v14w30 2→5：tool=182 构型下 ~5mm 固有误差映射关节达 2.58°（10-21 P8 实证），阈外即误判未执行——粗验收前哨放宽，法兰级粗验收(≤8mm/≤1°)+MoveJ收口紧随其后罩终点；此处不走 MOVE_OFFSET_TOL=0.5°（require_joints=False 路径，护栏语义不降级）

# v14w22：实机关节限位（与 RoboDK 模型 ±360 取交集）。依据：J1=193.59 两次被控制器
# -40001 拒收（10-15 P25）；J6=190.84 return 0 ✓；J5=177.6 实机走成 ✓（故 J5=180 非
# 某些资料的 ±120）；J3 取模型更紧的 ±160。规划期过滤，保证预检路径=实发路径。
# v14w23：J4 190→150——J4=-189.70 被控制器 -40004（自干涉 PoseSelfInterference）拒收；
# -168 族中途自干涉保护停机；实证安全族 |J4|≤95，150 留 55° 余量。
# ★★★ 2026-11-03：J4 150→178（用户要求）★★★
#   原因：150 太紧 ⇒ 某些点的【全部 IK 解都被过滤】⇒ 报 "ValueError: 没有限位内的逆解"
#         （11-03 10:29:35 实测：已完成 0 点即停）。要让那些点出解，J4 必须 ≥165。
#   代价：(150,178] 区间【重新暴露 -40004 自干涉拒收】风险 ✗
#         ⇒ 依靠 REAL_INTERFERE_J4_MAX / REAL_INTERFERE_J5_MIN（J4×J5 组合区禁选）
#           + 规划期预检（MoveJ_Test / MoveL_Test）兜底；
#         ⇒ 若再现 -40004，把本值在 165~178 之间微调（165 = "能出解 + 少踩禁区"的折中）。
#   历史：190 ✗(-40004) → 150 ✓（安全但出解困难）→ 178（本次，兼顾出解）
REAL_JOINT_LIMITS = (180.0, 180.0, 160.0, 178.0, 180.0, 360.0)

# v14w26：实机自干涉组合区（控制器 PoseSelfInterference 的 J4×J5 耦合，-40006）。
# 实录：|J4|=115.5×|J5|=173.1 与 |J4|=109.4×|J5|=171.5 均拒；|J4|=83.2×|J5|=177.6 通过。
# 阈值取中：|J4|>100 且 |J5|>165 视为禁区（两端各留 ~9°/~8° 实证余量）。
REAL_INTERFERE_J4_MAX = 100.0
REAL_INTERFERE_J5_MIN = 165.0
# ★★★ v15.2（2026-11-03）：【J4 单独硬禁区 |J4|>150】
#   背景：v15 把 J4 限位 150→178 之后，P5 的规划解从 J4=123.60° 变成 J4=172.88°（11-03 11:14:37 实录），
#         ⇒ 实机报「断连收尾后未到位…173.19…误差0.84°」，界面显示姿态自干涉 ✗（= 用户说的"原本没有的自干涉"）
#   现有组合禁区 (|J4|>100 且 |J5|>165) 抓不住它：P5 的 J5 只有 58.81° ⇒ 不在禁区 ⇒ 放行 ⇒ 踩雷 ✗
#   ⇒ 新增：|J4| > 150 一律视为禁区（与 v14w23 的"实证安全族 |J4|≤95、150 留 55° 余量"一致）
#   ⇒ 效果：J4 限位仍是 178（能出解、不误杀"没有限位内的逆解"），但【选中的解 J4 必 ≤150】
#          ⇒ P5 回到 J4=123.60 的原解 ⇒ 既出解又不自干涉 ✓
REAL_INTERFERE_J4_HARD = 150.0


def _real_interfere_combo(q):
    """v14w26：关节是否落入实机自干涉组合禁区（J4×J5 耦合，控制器 -40006）。
    v15.2：追加 |J4|>150 的单独硬禁区（治 P5 的 J4=172.88 自干涉）。"""
    if abs(q[3]) > REAL_INTERFERE_J4_HARD:
        return True
    return abs(q[3]) > REAL_INTERFERE_J4_MAX and abs(q[4]) > REAL_INTERFERE_J5_MIN


def _real_limit_ok(q, lower, upper):
    """v14w22：关节目标是否同时满足模型限位与实机限位。"""
    for j in range(min(6, len(q))):
        lo = max(float(lower[j]), -REAL_JOINT_LIMITS[j])
        hi = min(float(upper[j]), REAL_JOINT_LIMITS[j])
        if not lo <= float(q[j]) <= hi:
            return False
    return True


def _try_set_tool_user():
    """Unsupported through this driver: RunCodeCustom becomes RunScript, not raw Tool/User."""
    raise ControllerMotionFault('当前驱动未验证Tool/User透传；禁止通过项目调用设置坐标系。')


def _movl_digit_safe_joints(q_target):
    """v14w：直发位姿数字净化 —— 控制器 MovL 参数校验 -30001 防御。

    实证（控制器 logs/all/log）：
      11:38:20 拒收 MovL(-0.000000,…,300.000000,90.000000,0.000000,-0.000000)
               → [MovL#820] the type of params is wrong: -30001
      15:55:51 接受 MovL(0.000000,…,299.999986,89.999995,-0.000003,0.000000) → return 0
    触发器（同目标、不同关节末位 ⇒ 不同参数形态 ⇒ 校验翻转）：
      x 负零/极小负 · rx 恰=+90.000000 · **三角(rx/ry/rz)负零——ry=-0 是 -30005 实锤**
      （10-15 09:16 与 10-14 拒收样本共同点；接受样本 ry 均为 +0）· rz=+180（保留防御）
      —— 同时设防，且只在零/边界区动手：
      · x ∈ (-0.01, 0.001) mm → 推到 ≥ +0.001（FK 位置与欧拉约定无关，可靠）
      · rx ∈ [89.999, 90.001] → 拉出该区（Pose_2_Fanuc 的 rx 与两份实录一致）
      · rz 为负零 (-0.0) → 推离
    手法：对发送关节贪心微扰（步长 0.0005°→0.05°，单关节累计 ≤0.05°，末端位移 ≲0.6mm
    ≪ 圆柱真裕度 19.9mm ≪ 法兰验收 8mm）；到位/法兰验收/MoveJ 收口仍对【原始认证关节】
    判定，收口回认证构型 —— 几何语义不变。P5 类非边界参数零扰动（首查即过，原样返回）。
    返回 (send_q, note)：无违规=(原关节,None)；成功=(微扰关节,说明)；失败=(None,原因)。"""
    def _digits(q):
        # v14w19：先按驱动下发格式（6位小数）定型再判——控制器校验的是字符串形态；
        # 客户端 Fanuc 与驱动在零点附近的正负号约定不一致，故三角一律推离零域。
        # v14w24：净化微扰可能把限位边界关节（如 J6=-360.00）推出模型限位，
        # SolveFK 会抛 TargetReachError——捕获后返回 None=不可行候选（评分置顶永不选中）。
        try:
            return [float('%.6f' % v) for v in Pose_2_Fanuc(robot.SolveFK(q))]
        except Exception:
            return None

    def _score(vals):
        if vals is None:
            return 1e9   # 越界候选：永不优于当前
        x, rx, ry, rz = vals[0], vals[3], vals[4], vals[5]
        s = 0.0
        if -0.01 < x < 0.001:                      # 零附近（含 -0.000000）且未达 +0.001
            s += (0.001 - x) / 0.001
        if 89.999 <= rx <= 90.001:                 # 恰卡 +90 边界（含 90.000000 整）
            s += (rx - 89.999) / 0.001
        # v14w19：三角必须整体离开零域 ≥0.001°——"-0.000000"形态是 -30005 实锤
        #（10-15 09:16/09:35 两次实录 ry 打印 -0.000000 均拒；-2e-7 打印即 -0.000000
        #  而浮点 !=0.0 会漏判；推离零域后客户端/驱动符号一致为正）
        for v in (rx, ry, rz):
            if abs(v) < 0.001:
                s += 1.0 + (0.001 - abs(v)) / 0.001
        if rz >= 179.999:                          # rz=+180 疑似越界（保留防御）
            s += 1.0 + (rz - 179.999) / 0.001
        return s

    base = list(q_target)
    cur = _score(_digits(base))
    if cur <= 0.0:
        return q_target, None
    q = list(base)
    solved = False
    for step in (0.0005, 0.002, 0.01, 0.05):
        improved = True
        while cur > 0.0 and improved:
            improved = False
            for j in range(6):
                for sgn in (1.0, -1.0):
                    q2 = q[:]
                    q2[j] += sgn * step
                    if abs(q2[j] - base[j]) > 0.05 + 1e-9:
                        continue
                    sc = _score(_digits(q2))
                    if sc < cur - 1e-12:
                        q, cur, improved = q2, sc, True
                        break
                if improved:
                    break
        if cur <= 0.0:
            solved = True
            break
    if not solved:
        return None, '发送位姿净化失败（边界参数 x/rx/rz 微调不出安全区）'
    touched = ['%s%+.4f' % ('J%d' % (k + 1), q[k] - base[k]) for k in range(6)
               if abs(q[k] - base[k]) > 1e-9]
    return q, '发送关节微扰 %s°（Δmax 对应末端 ≪1mm）：规避 -30001 边界参数；验收/收口仍回认证构型' \
        % ' '.join(touched)


def _movl_flange_accept(joints_now, joints_target):
    """v14q：直发 MovL 落点的法兰位姿级粗验收。

    v14p 首航实证：控制器 MovL 固有落点残差 ~5mm/0.6° 级（v14p 4.61mm/0.616°、v14l 5.5mm，
    双样本跨版本一致）——关节级 0.5° 判据会把正常落点误判为事故。改用法兰语义验收：
    FK(实测) vs FK(目标)，位置≤MOVL_FLANGE_TOL_MM 且姿态≤MOVL_FLANGE_TOL_DEG 即过；
    过后在 _execute_checked_real 里发一条 MoveJ 微纠偏收口（关节级 0.5° 校验罩住终点）。
    超容差=落点异常（构型翻转/卡住/送错目标），照旧抛 RuntimeError 即停待判读。"""
    _f_now = invH(robot.PoseFrame()) * robot.SolveFK(joints_now)      # 法兰位姿（无工具）
    _f_tgt = invH(robot.PoseFrame()) * robot.SolveFK(joints_target)
    _d = _f_now * invH(_f_tgt)
    _mm = norm(_d.Pos())
    _deg = math.degrees(pose_angle(_d))
    return _mm, _deg


def _movl_direct_ready():
    """v14p 法兰补偿MOVL 开关是否可用：GUI 变量已建（正常运行）才开；
    离线 verify 的 exec 命名空间里没有 real_movldirect_var（NameError），
    自动回 False——离线验证的计划/指纹与该开关无关（规划层零改动）。"""
    try:
        return isinstance(real_movldirect_var, tk.BooleanVar)
    except Exception:
        return False


MOVE_SEGMENT_MAX_DEG = 64.0  # 每瓣最大关节跨度：驱动约8秒无完成回报即断连，20°/s下64°≈3秒，留足裕量


J6_SPIN_SEGMENT_DEG = 60.0   # MoveL 纯J6自转段分瓣跨度（无平移时关节插值=笛卡尔路径）


def _is_pure_j6_spin(start, target):
    """MoveL 目标仅 J6 变化（J1~J5 不动）：关节插值与笛卡尔路径重合，可精确分瓣。"""
    return max(abs(a - b) for a, b in zip(start[:5], target[:5])) < 1e-6


def _move_with_completion_check(method, target, allow_split=True):
    """长运动分瓣执行（v9）：驱动对单条指令约8秒无完成回报就断连（本环境常态，
    test.py 同款假报，它每段部在几秒内完成所以从没撞上）；大跨度关节运动沿
    预检验证过的同一条关节直线剖成若干瓣，每瓣都在死线内完成，路径不变，
    仅增设停顿点。MoveL 纯J6自转段同理分瓣；带平移 MoveL 与小跨度段保持原样。"""
    if not allow_split:
        # v11: 单点运动/关节运动不分瓣，恢复一指令直达（到位校验与假断连容忍保留）
        _single_move_settle(method, target)
        return
    try:
        start = _live_joints()
        total = max(abs(float(b) - float(a)) for a, b in zip(start, target))
    except Exception:
        start, total = None, None
    if method == 'MoveJ' and total is not None and total > MOVE_SEGMENT_MAX_DEG:
        pieces = int(math.ceil(total / MOVE_SEGMENT_MAX_DEG))
        log('长运动分瓣：跨度%.1f° → %d 瓣执行（同一关节直线，仅增设停顿点）。' % (total, pieces))
        for k in range(1, pieces + 1):
            way = [a + (b - a) * k / pieces for a, b in zip(start, target)]
            _single_move_settle('MoveJ', way)
            _require_joints(way)  # 瓣间校验到位，也给驱动链路留出响应时间
        return
    if (method == 'MoveL' and total is not None and _is_pure_j6_spin(start, target)
            and total > J6_SPIN_SEGMENT_DEG):
        pieces = int(math.ceil(total / J6_SPIN_SEGMENT_DEG))
        log('J6自转分段：跨度%.1f° → %d 段MoveL（纯自转，路径与笛卡尔路径重合）。' % (total, pieces))
        for k in range(1, pieces + 1):
            way = [a + (b - a) * k / pieces for a, b in zip(start, target)]
            _single_move_settle('MoveL', way)
            _require_joints(way)
        return
    _single_move_settle(method, target)


_real_running = False  # 2026-10-09 补回：旧版 L510 有此初始化，升级版漏带导致点击即 NameError 静默炸裂


def _ensure_canonical_tool():
    """v14w17：工具坐标守护——检测到 identity(0)（存档僵尸/直发残留）自动恢复规范值并大声记日志。
    实发两次：2026-10-14 18:2x、2026-10-15 09:0x（归零→种子/P2 预检异常、P5 直发异常）。
    v14w39：同时恢复被直发窗口残留隐藏的门把手（GUI 中途被杀会留下隐藏态→预检漏检）。
    每次执行入口 + 程序启动各调一次；非零值不干预（可能正在被人工调整）。"""
    if _tool_window_depth:
        return False  # Do not undo the intentional identity TCP during MOVL.
    pose = robot.PoseTool()
    fixed = False
    canonical = Fanuc_2_Pose(list(CANONICAL_TOOL))
    if _same_tool_pose(pose, eye(4)) or _same_tool_pose(pose, canonical):
        tcp = _named_tool(TCP_TOOL_NAME, canonical)
        _restore_tool(canonical, tcp)
    if _same_tool_pose(pose, eye(4)):
        log('⚠️ 工具坐标为0（存档残留/直发残留）——已自动恢复 [0,0,130]，请确认后再跑。')
        fixed = True
    try:
        _gh = RDK.Item('门把手_bs1')
        if _gh.Valid() and not _gh.Visible():
            _gh.setVisible(True)
            log('⚠️ 门把手网格处于隐藏态（直发窗口残留）——已恢复显示。')
            fixed = True
    except Exception:
        pass
    return fixed


def _execute_checked_real(data, single_method=None):
    global _real_running
    log('【入口】_execute_checked_real：%d 点，single_method=%s' % (len(data) if data is not None else -1, single_method))
    if _real_running:
        log('已有实机任务正在执行。')
        return
    _real_running = True
    completed = 0
    movl_direct = False  # v14p：入口预置，防异常早于赋值时 except 块二次 NameError（v14l 教训）
    try:
        _ensure_canonical_tool()  # Failure must pass through task cleanup.
        log('开始校验录入数据…')
        records = _validated_records(data)
        log('录入数据校验通过：%d 点。' % len(records))
        if single_method is None and len(records) > 1:
            expanded = _retreat_orientation_records(records)
            log('连续轨迹：%d个录入点展开为%d个执行点（含姿态退让）。' % (len(records), len(expanded)))
            records = expanded
        deviation = float(real_deviation_var.get())
        if not math.isfinite(deviation) or deviation < 0:
            raise ValueError('允许偏离必须为非负有限数。')
        log('偏离上限 %.1f mm，检查机器人连接…' % deviation)
        if not ensure_connected():
            return
        start = _live_joints()
        log('实机当前关节：%s' % ['%.2f' % v for v in start])
        # 长预检/运动期间 RoboDK 主程序忙或不消费驱动输出，驱动链路会饿死断开（15:20:56 P1 中途断连同因）。
        # 保活线程用独立 API 连接（避免被 MoveJ 阻塞主连接），每2秒一次 ConnectedState（只读），
        # 贯穿预检+执行全程，直到任务结束才停（v7 错在预检后就停，P1 运动中饿死驱动）。
        import threading as _th
        _keepalive_stop = _th.Event()
        def _driver_keepalive():
            n = 0
            _ka_rdk = Robolink()
            _ka_robot = _ka_rdk.Item(robot.Name(), ITEM_TYPE_ROBOT)
            while not _keepalive_stop.wait(2.0):
                n += 1
                try:
                    s, _m = _ka_robot.ConnectedState()
                    if s < 0:
                        log('【保活】第%d次发现驱动掉线（%s），已请求重连。' % (n, _m))
                        _ka_robot.Connect()
                except Exception:
                    pass  # 主程序忙时 API 调用可能慢/超时，下一轮再试
        _ka_thread = _th.Thread(target=_driver_keepalive, daemon=True, name='driver_keepalive')
        _ka_thread.start()
        log('已启驱动保活（贯穿预检+执行）。')
        frame, tool = robot.PoseFrame(), robot.PoseTool()
        log('开始台子/地面避障预检，尚未发送运动指令。')
        plan = _prepare_real_plan(records, start, deviation, single_method)
        # 保活线程不在此处停：执行阶段同样需要（v7 教训）
        # 预检后复核：驱动必须就绪且关节与预检起始一致，否则取消。
        if not ensure_connected():
            log('预检后驱动断连，重连未成功，取消执行。')
            return
        _require_joints(start)
        log('预检后连接复核通过，准备发运动指令。')
        # v14w22：实机限位最后防线（规划器已过滤，此处兜底拦截任何漏网目标）
        # ★ v15（2026-11-03）：判限位前先做【同角归一化】—— 修一次误拦：
        #   实录 11:07:59 `段6 目标关节超出实机限位：['64.99','77.69','-96.48','198.78','64.99','0.00']`
        #   而 198.78° 与 −161.22° 是【同一个角】（差 360°），规划期用的是 −161.22（合法 ✓），
        #   最后防线却拿 198.78 去比 ⇒ 误判超限 ⇒ 整段 0 点即停 ✗。
        #   ⇒ 对每个关节先试 ±360k 的等价表示，取限位内的那个；都不在限位内才判死。
        #   ⇒ 并把归一化后的值【写回 plan】，避免执行时把 198.78 发给控制器（J6 合法域 ±360，故按轴各自限位判）。
        _lo, _hi, _ = robot.JointLimits()
        _lo, _hi = _lo.list(), _hi.list()

        def _nearest_in_limit(q):
            out = []
            for j in range(6):
                v = float(q[j])
                lo = max(float(_lo[j]), -REAL_JOINT_LIMITS[j])
                hi = min(float(_hi[j]), REAL_JOINT_LIMITS[j])
                if lo <= v <= hi:
                    out.append(v)
                    continue
                picked = None
                for k in (-1.0, 1.0):
                    alt = v + 360.0 * k
                    if lo <= alt <= hi:
                        picked = alt
                        break
                out.append(picked if picked is not None else v)
            return out

        for _i, _step in enumerate(plan, 1):
            _q_raw = list(_step['joints'])
            _q_near = _nearest_in_limit(_q_raw)
            if _q_near != _q_raw:
                log('段%d 关节取同角等价表示：%s → %s'
                    % (_i, ['%.2f' % v for v in _q_raw], ['%.2f' % v for v in _q_near]))
                _step['joints'] = _q_near[:]          # 执行也用归一化值 ✓
            if not _real_limit_ok(_step['joints'], _lo, _hi):
                raise ValueError('段%d 目标关节超出实机限位：%s（规划期应已过滤，此为最后防线；已试 ±360 同角表示）'
                                 % (_i, ['%.2f' % v for v in _step['joints']]))
        for before, after in ((frame, robot.PoseFrame()), (tool, robot.PoseTool())):
            error = invH(before)*after
            if norm(error.Pos()) > 0.01 or pose_angle(error) > math.radians(0.01):
                raise RuntimeError('预检期间工具或参考坐标系改变，取消执行。')
        robot.setSpeed(ROBOT_SPEED)
        RDK.Command('Trace','Reset')
        RDK.Command('Trace','On')
        expected = start
        # v14k：停用长运动分瓣（split_moves 恒 False）。2026-10-12 实测日志坐实：假断连与跨度无关，
        # 60°/95°/169°/180° 的瓣与 20mm 途经点每条指令都在断，分瓣已不防任何东西，只剩每瓣一轮
        # 等待+重连停顿税；_single_move_settle 断连容忍（_wait_controller_static 20s 静止上限）
        # 罩得住单条长指令的收尾（20°/s 下 180°≈9s<20s）。分瓣机制与常量原样留档，遇真断连指纹
        # （未自然收尾/未到位）随时把本行改回 single_method is None and len(records) > 1 即可恢复。
        split_moves = False
        movl_direct = bool(real_movldirect_var.get()) if _movl_direct_ready() else False
        if movl_direct:
            # v15：原来的超长版本横幅已按用户要求删除，只留一行关键参数，便于判读
            log('直发开启 ｜ 段长≤%.0fmm ｜ 法兰容差 %.0fmm/%.1f° ｜ 等待≤%.0fs ｜ 禁直发名单=%s'
                % (MOVL_DIRECT_MAX_MM, MOVL_FLANGE_TOL_MM, MOVL_FLANGE_TOL_DEG,
                   MOVL_ARRIVE_WAIT_S, MOVL_DIRECT_BLOCK_POINTS))
        log('本次单条MovL动态认证放行点=%s' % [i for i,s in enumerate(plan,1) if s.get('direct_movl_certified')])
        _assert_continuous_dispatch(records, start, plan, movl_direct)
        for i, step in enumerate(plan, 1):
            for rewind in step['rewinds']:
                _require_joints(expected)
                _move_with_completion_check("MoveJ", rewind, split_moves)
                _require_joints(rewind)
                expected = rewind
            _require_joints(expected)
            waypoints = step.get('waypoints') or []
            if step['method'] == 'MoveL' and not waypoints:
                # 理论不可达：v13 起所有 MoveL 步都带细分途经点；不带则说明规划层契约被破坏
                raise RuntimeError(f"P{i}：MoveL 步缺少细分途经点，拒绝发送驱动 MOVL（已判死）。")
            seg_mm = seg_rot = None
            if movl_direct and step['method'] == 'MoveL' and waypoints:
                # 仅开关开启时才算（两次 FK 的 API 往返）；开关关/离线 verify 零开销
                _seg_rel = _trajectory_pose(step['joints']) * invH(_trajectory_pose(expected))
                seg_mm, seg_rot = norm(_seg_rel.Pos()), pose_angle(_seg_rel)
            direct_ready = (movl_direct and _direct_step_allowed(i, step)
                            and seg_mm is not None
                            and seg_mm <= MOVL_DIRECT_MAX_MM
                            and seg_rot <= math.radians(0.5))
            _send_q = step.get('direct_send_joints', step['joints'])
            if direct_ready and not step.get('direct_movl_certified'):
                # v14w：发送前数字净化——控制器 -30001 拒的是【参数形态】不是几何（LOG_VERSION
                # 处 11:38 拒收 / 15:55 接受两份实录）。净化只在零边界区微调发送关节；
                # 净化失败 ⇒ direct_ready=False ⇒ 落到 elif waypoints 走细分（安全回落）。
                _send_q, _purge_note = _movl_digit_safe_joints(step['joints'])
                if _send_q is None:
                    log('P%d：⛔ %s ⇒ 改走细分途经点路径。' % (i, _purge_note))
                    direct_ready = False
                elif _purge_note:
                    log('P%d：%s' % (i, _purge_note))
            if direct_ready:
                # v14p 法兰补偿MOVL：驱动 MOVL 无工具补偿、按法兰执行（v14l 11:30 实证停点法兰=
                # 命令TCP目标，差仅5.5mm）——将错就错：把本步构型的【法兰位姿】直接当笛卡尔目标
                # 发给控制器，法兰被精确送到位，物理工具尖端（182mm，v14w27 实测）随之落在认证
                # 直线上。姿态恒定段法兰线=TCP线平移常向量，扫掠包络与细分路径一致。
                # v14w36/37 演进：v14w36 只改传位姿（不切工具）⇒ MoveL(位姿) 按 TCP 空间
                # 校验，P8 法兰位姿被反推到 z=744 爆臂展 TargetReachError（11:18 实录）；
                # v14w37 = 位姿传递（动画=认证直线，根治关节弧假碰撞冻死）+ 发送窗口单位
                # 变换（校验/数字=法兰空间）；柜子实收参数与旧金标准逐位一致（0 偏差）。
                log(f"P{i}：v14w 法兰补偿MOVL：段长{seg_mm:.1f}mm（姿态变化{math.degrees(seg_rot):.2f}°），收起 {len(waypoints)} 个细分途经点，一指令直发（发法兰位姿=自算FK+单位变换窗口，发送关节已净化；v14w37）。")
                # v14r：require_joints=False——假断连分支的关节级 0.5° 校验让位给下方
                # 法兰级粗验收+MoveJ 微纠偏收口（终点仍回认证构型，护栏语义不降级）。
                # v14u：expect_target=段目标关节——目标锚定到位等待（上限 60s，每5s进度日志）。
                # v14w：净化只作用于发送关节；expect_target 仍是认证关节（到位判据不变）。
                # v14w37：位姿传递（动画=认证直线）+ flange_space 单位变换（校验/数字=法兰空间）。
                _send_pose = invH(robot.PoseFrame()) * robot.SolveFK(_send_q)
                # ★ 2026-11-03（可选，默认关）：先给控制器发 Tool(0)/User(0)，
                # 治 `[MovL#878] movL not set tool or user!!!` ⇒ 让 MovL 明确按 基座系+零工具(法兰) 执行。
                # 打开方式：把 MOVL_SEND_TOOL_USER 改成 True（建议先跑一条短段验证）。
                if MOVL_SEND_TOOL_USER:
                    if _try_set_tool_user():
                        log('  ✓ Tool(0)/User(0) 已下发，继续直发')
                    else:
                        raise ControllerMotionFault('Tool/User未确认，停止直发。')
                log('P%d：发送法兰目标=%s；认证关节=%s；TCP=%s' % (i, Pose_2_Fanuc(_send_pose), step['joints'], Pose_2_Fanuc(robot.PoseTool())))
                _single_move_settle('MoveL', _send_pose, require_joints=False,
                                    expect_target=step['joints'], flange_space=True)
                # ★★★ v15.7（2026-11-03）：直发结束后【先等真静止】再做后续（法兰验收/收口）。
                #   实录（v15.6, P8）：直发报"已完成"（假断连分支）→ 脚本立刻法兰验收(5.71mm ✓)
                #   → P8 尾部关节检查【通过】（读到的是过渡中姿态）→ P9 开头再读【已翻转】⇒ 差 20~38° ⇒ 停 ✗
                #   对比：P7 目标 [75.42,12.24,57.74,20.02] vs 停止实测 [78.10,36.86,19.48,33.66]
                #         ⇒ J2↑25 / J3↓38 / J4↑14 = 典型【肘部翻转 elbow flip】✗
                #   机理：MovL 只给位姿 ⇒ 控制器自行选 IK 分支（可能选翻转那组）✗
                #         + 直发"已完成"没等真静止 ⇒ 后续读到的是过渡值 ✗
                #   ⇒ 这里补一段【关节稳定等待】：连续 3 次采样（每次 0.3s）关节变化 <0.05° 才算真停，
                #     最多等 8 秒；等稳定后再做验收/收口，避免"读到过渡值"造成的假通过/假失败。
                _st = None
                _stable = False
                for _w in range(24):          # 24 × 0.3s ≈ 7.2s 上限
                    _cur = _live_joints()
                    if _st is not None and max(abs(a - b) for a, b in zip(_cur, _st)) < 0.05:
                        _stable = True
                        break
                    _st = _cur
                    time.sleep(0.3)
                if not _stable:
                    log('P%d：⚠️ 直发后 7 秒内关节仍未稳定（继续按现值验收，可能判死）' % i)
                else:
                    log('P%d：直发后关节已稳定 ✓（进入法兰验收/收口）' % i)
                # ★★★ v15.8（2026-11-03）：★ 安全网 —— 直发是【控制器自行选 IK 解】，
                #   规划期的自干涉硬禁区（|J4|>150 等）拦不到它 ✗
                #   ⇒ 直发落点若真落进禁区（J4 极端 / J4×J5 组合区），必须【立刻回认证构型】，
                #     绝不能把手臂留在危险姿态里继续跑下一段 ✓
                _post = _live_joints()
                if _real_interfere_combo(_post):
                    log('P%d：🚨 直发落点落入自干涉禁区！实测=%s（J4=%.2f J5=%.2f）⇒ 立即回认证构型'
                        % (i, ['%.2f' % v for v in _post], _post[3], _post[4]))
                    _single_move_settle('MoveJ', step['joints'])
                    _require_joints(step['joints'])
                    log('P%d：已回到认证构型 ✓' % i)
                elif abs(_post[3]) > REAL_INTERFERE_J4_MAX:
                    log('P%d：⚠️ 直发落点 J4=%.2f° 偏大（>%.0f° 组合区阈值，但未触禁区组合）——记录'
                        % (i, _post[3], REAL_INTERFERE_J4_MAX))
                try:
                    robot.setJoints(_post)   # 显示实测姿态，不用预期目标掩盖未到位。
                except Exception:
                    pass
                # v14q：MovL 落点法兰级粗验收（≤8mm/≤1°）+ MoveJ 微纠偏收口（关节级 0.5° 罩终点）。
                # v14p 首航停在 0.95° 关节残差（法兰 4.61mm/0.616°）被 0.5° 护栏拦停——那是控制器
                # MovL 固有落点残差（v14l 5.5mm 双样本背书），不是构型错误；但终点必须回到认证构型，
                # 故验收通过后用一条短 MoveJ（~1° 关节差）收口，走 _single_move_settle 全套护栏。
                _actual, _is_static = _wait_controller_static(samples=3, interval=0.2)
                _mm, _deg = _movl_flange_accept(_actual, step['joints'])
                if _mm > MOVL_FLANGE_TOL_MM or _deg > MOVL_FLANGE_TOL_DEG:
                    raise RuntimeError('v14u 法兰级粗验收未过：停点法兰残差%.2fmm/%.2f°（容差%.1fmm/%.1f°），实测关节%s，停止待判读。'
                                       % (_mm, _deg, MOVL_FLANGE_TOL_MM, MOVL_FLANGE_TOL_DEG,
                                          ['%.2f' % v for v in _actual]))
                _jm = max(abs(a - b) for a, b in zip(_actual, step['joints']))
                if _jm > MOVE_OFFSET_TOL:
                    log(f"P{i}：v14u MovL 直发落点法兰级验收通过（残差{_mm:.2f}mm/{_deg:.2f}°），关节残差{_jm:.2f}°——发 MoveJ 微纠偏收口。")
                    # ★★★ v15.4（2026-11-03）：收口 MoveJ 加重试 —— 治"P8 停下"：
                    #   实录 11:29:03 验收通过 → 发收口 MoveJ → 11:29:04 驱动报断连 → 11:29:06 才重连
                    #   ⇒ 那条收口 MoveJ 没走完 ⇒ 关节残差 2.68° 残留
                    #   ⇒ 下一段前的 _require_joints（容差 0.5°）判死 ⇒ 停在 P8 ✗
                    #   收口目标是【认证构型】（确定可达）⇒ 重发安全 ✓；最多 2 次，仍不到就抛原错。
                    _close_err = None
                    for _close_try in (1, 2):
                        try:
                            _single_move_settle('MoveJ', step['joints'])
                            _close_err = None
                            break
                        except Exception as _close_exc:  # noqa: BLE001
                            _close_err = _close_exc
                            if _close_try == 1:
                                log('P%d：收口 MoveJ 未完成（%s: %s）⇒ 重试一次（目标为认证构型，可达）'
                                    % (i, type(_close_exc).__name__, _close_exc))
                                time.sleep(0.5)
                    if _close_err is not None:
                        raise _close_err
                # ★★★ v15.5（2026-11-03）：直发+收口之后，再做【关节校正重试】—— 治 P8 停下的真因。
                #   实录（v15.4, 11:36:19~23）：
                #     P8 直发到位（关节残差 2.68°）→ 法兰验收通过 → 发收口 MoveJ
                #     → 驱动报断连 → 脚本打印「驱动断连但运动已自然完成到位」（★ 它认为完成 ✗）
                #     → 于是 _single_move_settle 没抛异常（断连分支 require_joints=False 不校验关节）
                #     → 紧接的 _require_joints 才发现不一致（实测 J2=36.86/J3=19.48，差很多）⇒ 抛错停 ✗
                #   ⇒ 所以 v15.4 的 try/except 重试【根本没触发】✗
                #   ⇒ 改为：_require_joints 失败时【再发一次定向 MoveJ】校正（目标=认证构型，确定可达）
                try:
                    _require_joints(step['joints'])
                except Exception:
                    log('P%d：直发+收口后关节仍与预检不一致 ⇒ 再发一次 MoveJ 校正（目标为认证构型，可达）' % i)
                    time.sleep(0.5)
                    _single_move_settle('MoveJ', step['joints'])
                    _require_joints(step['joints'])
                    log('P%d：校正 MoveJ 完成 ✓' % i)
            elif (movl_direct and not _direct_step_allowed(i, step) and seg_mm is not None
                    and seg_mm <= MOVL_DIRECT_MAX_MM and seg_rot <= math.radians(0.5)):
                # ★ v14v4：本点被【禁直发名单】拦下 —— 明确告知，便于判读日志
                log(f"P{i}：⛔ 本点在【禁直发名单】MOVL_DIRECT_BLOCK_POINTS={MOVL_DIRECT_BLOCK_POINTS} 里 ⇒ "
                    f"不走法兰补偿直发，改走【细分途经点路径】（v14n 实测 17/17 通过、零事故的路径）。")
                if not waypoints:
                    raise RuntimeError(f'P{i}：禁直发点缺少途经点，停止。')
                for way in waypoints:
                    _move_with_completion_check('MoveJ', way, False)
                    _require_joints(way)
                _require_joints(step['joints'])
            elif waypoints:
                log(f"P{i}：执行预检方案 {step['method']}→MoveJ 细分，{len(waypoints)} 个途经点，终点关节={step['joints']}")
                for k, way in enumerate(waypoints, 1):
                    _move_with_completion_check('MoveJ', way, False)
                    _require_joints(way)
                _require_joints(step['joints'])
            else:
                log(f"P{i}：执行预检方案 {step['method']}，关节={step['joints']}")
                _move_with_completion_check(step['method'], step['joints'], split_moves)
                _require_joints(step['joints'])
            expected = step['joints']
            completed += 1
        log(f'实机执行完成：{completed}/{len(plan)}点。')
    except Exception as exc:
        log(f'实机任务停止，已完成{completed}点：{type(exc).__name__}: {exc}')
        if movl_direct and ('断连' in str(exc) or '未到位' in str(exc) or '落点偏差' in str(exc) or '粗验收' in str(exc)):
            log('【v14u】法兰补偿MOVL执行段出断连/落点指纹（v14w24 无勾选框；细分途经点路径保留在计划中，可作回退依据）。')
        try:
            actual, velocity, mode = _controller_feedback()
            log('停止时控制器实际反馈：关节=%s，速度=%s，模式=%s；不自动重发运动。' % (actual, velocity, mode))
        except Exception as feedback_error:
            log('停止时也无法取得控制器反馈：%s' % feedback_error)
    finally:
        _real_running = False
        try:
            _keepalive_stop.set()
            _ka_thread.join(timeout=3)
        except Exception:
            pass


def _point_to_segment_distance(p, a, b):
    """3D点到线段距离，单位mm。"""
    ax, ay, az = a
    bx, by, bz = b
    px, py, pz = p
    ab = (bx-ax, by-ay, bz-az)
    ap = (px-ax, py-ay, pz-az)
    ab2 = ab[0]*ab[0] + ab[1]*ab[1] + ab[2]*ab[2]
    if ab2 < 1e-12:
        return math.sqrt((px-ax)**2 + (py-ay)**2 + (pz-az)**2)
    t = (ap[0]*ab[0] + ap[1]*ab[1] + ap[2]*ab[2]) / ab2
    t = max(0.0, min(1.0, t))
    q = (ax+t*ab[0], ay+t*ab[1], az+t*ab[2])
    return math.sqrt((px-q[0])**2 + (py-q[1])**2 + (pz-q[2])**2)


def _tcp_position_from_joints(q):
    """关节角 -> 当前参考坐标系下的TCP位置，与轨迹输入使用同一坐标系。"""
    f = pose_to_fanuc_values(invH(robot.PoseFrame()) * robot.SolveFK(q) * robot.PoseTool())
    return (float(f[0]), float(f[1]), float(f[2]))


def _check_movej_tcp_trajectory(start_q, target_q, start_tcp_vals, target_tcp_vals, log, samples=30, max_deviation_mm=None):
    """
    在真正执行MoveJ之前，用关节空间线性插补采样，计算TCP轨迹相对
    起点-终点TCP直线段的最大偏离距离。

    目的：MoveL失败时，不再无条件MoveJ；只有MoveJ造成的TCP空间绕行
    没有超过允许值，才允许用MoveJ兜底。
    """
    if max_deviation_mm is None:
        max_deviation_mm = MOVEJ_FALLBACK_MAX_DEVIATION_MM

    start_q = [float(v) for v in start_q[:6]]
    target_q = [float(v) for v in target_q[:6]]
    a = (float(start_tcp_vals[0]), float(start_tcp_vals[1]), float(start_tcp_vals[2]))
    b = (float(target_tcp_vals[0]), float(target_tcp_vals[1]), float(target_tcp_vals[2]))

    log("开始检查 MoveJ 兜底轨迹：%d 个采样点，允许最大TCP偏离 %.3f mm" % (samples + 1, max_deviation_mm))
    max_dev = -1.0
    max_info = None

    for k in range(samples + 1):
        t = float(k) / float(samples)
        q = [start_q[j] + (target_q[j] - start_q[j]) * t for j in range(6)]
        try:
            p = _tcp_position_from_joints(q)
        except Exception as e:
            log("  MoveJ轨迹检查失败：第 %d/%d 个采样点 FK失败：%s: %s" % (k+1, samples+1, type(e).__name__, e))
            return False

        dev = _point_to_segment_distance(p, a, b)
        if dev > max_dev:
            max_dev = dev
            max_info = (k, t, q, p)

        if dev > max_deviation_mm:
            log("✕ MoveJ兜底轨迹拒绝：第 %d/%d 个采样点偏离TCP直线 %.3f mm > %.3f mm" %
                (k+1, samples+1, dev, max_deviation_mm))
            log("  t=%.3f  TCP=(%.3f, %.3f, %.3f)" % (t, p[0], p[1], p[2]))
            log("  因此不会执行这个MoveJ兜底动作，避免出现不可接受的大绕圈。")
            return False

    if max_info is not None:
        k, t, q, p = max_info
        log("✓ MoveJ兜底轨迹检查通过")
        log("  最大TCP偏离直线：%.3f mm（采样 %d/%d，t=%.3f）" % (max_dev, k+1, samples+1, t))
        log("  最大偏离点TCP=(%.3f, %.3f, %.3f)" % (p[0], p[1], p[2]))
    return True


# ============================================================
# 执行连续运动（MoveL失败时先检查MoveJ轨迹）
# ============================================================
def _collision_details():
    pairs = RDK.CollisionPairs()
    return '；'.join(f'{a.Name()}[连杆{ia}] 与 {b.Name()}[连杆{ib}]'
                    for a, b, ia, ib in pairs) or '路径碰撞或关节不可行'


def _enable_obstacle_checks():
    if RDK.RunMode() != RUNMODE_SIMULATE:
        raise RuntimeError('障碍物预检仅允许在仿真模式执行。')
    # 每次进入预检都清空预检缓存：缓存生命周期 = 单次预检规划，
    # 障碍物/工作站状态的变化在下一次预检即时生效。
    _plan_cache.clear()
    for name in ('安装台_650x650x80mm', '地面_禁止穿越', '磨砂圆柱_R150_H50', '挡板_半封闭3面'):
        obstacle = RDK.Item(name, ITEM_TYPE_OBJECT)
        if not obstacle.Valid():
            raise RuntimeError(f'缺少障碍物模型：{name}，请加载包含台子和地面的工作站。')
        if name == '安装台_650x650x80mm':
            if RDK.setCollisionActivePair(COLLISION_OFF, robot, obstacle, 0, 0) != 1:
                raise RuntimeError('无法配置安装台与固定底座的接触关系。')
        for link in range(1, 7):
            if RDK.setCollisionActivePair(COLLISION_ON, robot, obstacle, link, 0) != 1:
                raise RuntimeError(f'无法启用{name}与连杆{link}的碰撞检查。')
        tool_items = list(RDK.ItemList(ITEM_TYPE_TOOL))
        _handle = RDK.Item('门把手_bs1')   # v14w12：网格替换后可能为 OBJECT 类型，按名并入
        if _handle.Valid() and all(_handle.item != t.item for t in tool_items):
            tool_items.append(_handle)
        for tool in tool_items:
            parent = tool.Parent()
            while parent.Valid() and parent.item != robot.item:
                parent = parent.Parent()
            if parent.Valid() and RDK.setCollisionActivePair(COLLISION_ON, tool, obstacle) != 1:
                raise RuntimeError(f'无法启用{name}与工具的碰撞检查。')
    RDK.setCollisionActive(COLLISION_ON)


def _check_single_joint_path(end):
    _enable_obstacle_checks()
    saved = robot.Joints().list()[:6]
    try:
        RDK.Command('Trace', 'Off')
        RDK.Render(False)
        if _movej_test_cached(saved, end, 1) != 0:
            raise ValueError('单点MoveJ路径被拒绝：' + _collision_details())
    finally:
        robot.setJoints(saved)
        RDK.Render(True)


def _trajectory_pose(q):
    return invH(robot.PoseFrame()) * robot.SolveFK(q) * robot.PoseTool()


def _reorient_next_pose(records, i, rec):
    """v14w33：i 为 1-based 点号。若下一点存在且为【同 TCP 位姿纯换姿】（xyz 全同、姿态不同），
    返回下一点的 TCP 位姿 Mat，否则 None。用于换姿对的分支前视。"""
    try:
        if i >= len(records):
            return None
        nxt = records[i]          # 0-based 列表：下一条记录
        if nxt['type'] != 'TCP' or nxt.get('singular', False):
            return None
        va = [float(v) for v in rec['values'][:6]]
        vb = [float(v) for v in nxt['values'][:6]]
        if all(abs(va[k] - vb[k]) < 1e-9 for k in range(3)) and any(abs(va[k] - vb[k]) > 1e-9 for k in range(3, 6)):
            return fanuc_values_to_pose(*vb)
    except Exception:
        return None
    return None


def _linear_path_endpoint(start, target):
    """带结果缓存：分支重试时同一（起点, 目标）不重复计算。"""
    key = ('linear', _cache_key_joints(start), _cache_key_pose(target))
    if key in _plan_cache:
        return _plan_cache[key]
    result = _linear_path_endpoint_uncached(start, target)
    _plan_cache[key] = result
    return result


def _linear_path_endpoint_uncached(start, target):
    # 粗筛：10mm 采样点是 1mm 采样点的子集，粗筛失败则 1mm 细查必然失败，
    # 可直接拒绝；粗筛通过后再跑原有 1mm 细查，通过/拒绝判定与只跑 1mm 完全一致。
    if RDK.RunMode() != RUNMODE_SIMULATE:
        raise RuntimeError('直线路径预检仅允许在仿真模式执行。')
    # v15.17: Lookahead may leave the model at the P10 wrist-spin posture.
    # RoboDK's numerical IK uses current model joints even with an explicit j1.
    # Reset the model seed before each independent path check.
    robot.setJoints(start)
    status = robot.MoveL_Test(start, target, minstep_mm=10)
    if status == 0:
        robot.setJoints(start)
        status = robot.MoveL_Test(start, target, minstep_mm=1)
    if status != 0:
        return None, f'MoveL原生路径检查未通过（{status}）：' + _collision_details()
    # 本机MoveL_Test返回成功后Joints()可能为全零；从插补矩阵读取实际终点。
    # 碰撞判定已由上方同路径 1mm MoveL_Test 完成，此处仅提取终点关节，
    # 关闭碰撞检查提速（实测约快两个数量级）；整段权威碰撞复核仍在
    # _verify_obstacle_plan（碰撞开、1mm）进行。
    program = RDK.AddProgram('_TCP仿真_路径预检', robot)
    try:
        program.setVisible(False)
        robot.setJoints(start)
        program.setPoseFrame(robot.PoseFrame())
        program.setPoseTool(robot.PoseTool())
        program.MoveJ(start)
        program.MoveL(target)
        message, matrix, status = program.InstructionListJoints(mm_step=1, deg_step=1, collision_check=COLLISION_OFF)
        if status < 0:
            return None, message
        end = matrix.tr().rows[-1][:6]
        error_pose = invH(target) * _trajectory_pose(end)
        if norm(error_pose.Pos()) > .01 or pose_angle(error_pose) > math.radians(.01):
            raise RuntimeError('路径预检返回的终点不匹配目标TCP。')
        return end, message
    finally:
        program.Delete()


def _linear_waypoints(start, target, step_mm=None):
    """v13：从一条 MoveL 指令采样细分途经关节点（按 IK 顺序，无分支翻转）。

    用 InstructionListJoints(mm_step=LINEAR_SUBSTEP_MM, collision_check=COLLISION_OFF) 采样：
    途经点与 MoveL 执行的是同一条几何直线，且 IK 连续选解（避免用全局 SolveIK 时
    途经点在多解间跳变）。碰撞已由 _linear_path_endpoint 的 MoveL_Test@1mm 权威判定，
    此处不再重复。返回含终点的关节点列表；空列表表示采样失败（调用方回退直达）。"""
    if step_mm is None:
        step_mm = LINEAR_SUBSTEP_MM
    key = ('waypoints', _cache_key_joints(start), _cache_key_pose(target), round(float(step_mm), 3))
    if key in _plan_cache:
        return [q[:] for q in _plan_cache[key]]
    program = RDK.AddProgram('_TCP仿真_细分采样', robot)
    saved = robot.Joints().list()[:6]
    try:
        program.setVisible(False)
        robot.setJoints(start)
        program.setPoseFrame(robot.PoseFrame())
        program.setPoseTool(robot.PoseTool())
        program.MoveJ(start)
        program.MoveL(target)
        message, matrix, status = program.InstructionListJoints(mm_step=step_mm, deg_step=1, collision_check=COLLISION_OFF)
        cols = matrix.tr().rows if matrix is not None else []
        if status < 0 or not cols:
            return []
        # 丢弃比步长更密的重复点（InstructionListJoints 在奇异附近会加密采样）
        picked = [list(map(float, cols[0][:6]))]
        for row in cols[1:]:
            q = list(map(float, row[:6]))
            if max(abs(a - b) for a, b in zip(q, picked[-1])) >= step_mm / 10.0:
                picked.append(q)
        # 去尾：InstructionListJoints 可能带比目标多一点的收尾点，以关节距离最近的为准
        end_q, _ = _linear_path_endpoint(start, target)
        if end_q is not None and picked and max(abs(a - b) for a, b in zip(end_q, picked[-1])) > 1.0:
            picked[-1] = list(map(float, end_q))
        _plan_cache[key] = [q[:] for q in picked]
        return [q[:] for q in picked]
    finally:
        program.Delete()
        robot.setJoints(saved)


def _obstacle_posture_key(q, reference=None):
    table = RDK.Item('安装台_650x650x80mm', ITEM_TYPE_OBJECT)
    height = 0.0
    if table.Valid():
        elbow = invH(table.PoseAbs()) * robot.PoseAbs() * robot.JointPoses(q)[3]
        height = elbow.Pos()[2]
    return (-round(height, 6), sum((v-r)**2 for v, r in zip(q, reference or [0]*6)), tuple(q))


def _obstacle_joint_target(start, values, max_deviation=None, log=None):
    """带结果缓存：同一（起点, 目标, 偏离上限）的兜底选解不重复搜索。"""
    key = ('obstacle', _cache_key_joints(start), tuple(round(float(v), 6) for v in values[:6]),
           round(float(max_deviation), 6) if max_deviation is not None else None)
    if key in _plan_cache:
        cached = _plan_cache[key]
        if isinstance(cached, ValueError):
            raise cached
        return cached
    try:
        result = _obstacle_joint_target_uncached(start, values, max_deviation, log)
    except ValueError as exc:
        _plan_cache[key] = exc
        raise
    _plan_cache[key] = result
    return result


def _obstacle_joint_target_uncached(start, values, max_deviation=None, log=None):
    # v14-P2P：不再用 seed 候选/肘高排序，直接取离当前关节最近的逆解做逐级检查；
    # 最近解过不了偏离/碰撞时仍会在这里报错（单点 MoveJ 兜底路径保持可用）。
    lower, upper, _ = robot.JointLimits()
    candidates = [_nearest_ik_from_current(start, fanuc_to_pose(*values))]
    saved = robot.Joints().list()[:6]
    try:
        # 少量FK采样仅用于排序；不能替代后面的偏离复核与精细碰撞检查。
        a = _tcp_position_from_joints(start)
        table = RDK.Item('安装台_650x650x80mm', ITEM_TYPE_OBJECT)
        base_to_table = invH(table.PoseAbs()) * robot.PoseAbs()
        ranked = []
        for end in candidates:
            deviation, height = 0.0, float('inf')
            for k in range(11):
                q = [x + (y-x)*k/10 for x, y in zip(start, end)]
                deviation = max(deviation, _point_to_segment_distance(
                    _tcp_position_from_joints(q), a, values[:3]))
                height = min(height, (base_to_table * robot.JointPoses(q)[3]).Pos()[2])
            if max_deviation is not None and deviation > max_deviation:
                continue
            # 20mm一档，避免为很小的偏离差反复搜索；同档优先抬高肘部。
            ranked.append(((int(deviation/20), -height,
                            sum(abs(y-x) for x, y in zip(start, end))), end))
        checked = 0
        for _, end in sorted(ranked, key=lambda entry: entry[0]):
            if max_deviation is not None and not _check_movej_tcp_trajectory(
                    start, end, pose_to_fanuc_values(_trajectory_pose(start)), values,
                    lambda msg: None, samples=100, max_deviation_mm=max_deviation):
                continue
            checked += 1
            if _movej_test_cached(start, end, .25) == 0:
                if log is not None:
                    log(f'MoveJ快速筛选：{len(candidates)}个候选，{len(ranked)}个通过粗筛，精查{checked}条后找到合格路径。')
                return end
        raise ValueError('所有候选关节路径均碰撞、超出偏离限制或没有有效逆解。')
    finally:
        robot.setJoints(saved)


def _verify_obstacle_plan(start, plan):
    program = RDK.AddProgram('_TCP仿真_整段碰撞复核', robot)
    saved = robot.Joints().list()[:6]
    try:
        program.setVisible(False)
        program.setPoseFrame(robot.PoseFrame())
        program.setPoseTool(robot.PoseTool())
        program.MoveJ(start)
        for step in plan:
            for q in step['rewinds']:
                program.MoveJ(q)
            if step['method'] == 'MoveL' and not step.get('waypoints'):
                # v13 防呆：MoveL 步必须带细分途经点，否则规划层契约被破坏
                raise ValueError('整段碰撞复核：MoveL 步缺少细分途经点，拒绝。')
            getattr(program, step['method'])(step['joints'])
        message, matrix, status = program.InstructionListJoints(
            mm_step=1, deg_step=1, collision_check=COLLISION_ON)
        if status < 0 or 'collision' in message.lower():
            raise ValueError('整段碰撞复核未通过：' + message)
    finally:
        program.Delete()
        robot.setJoints(saved)


# Continuous TCP paths always recover calibrated-body IK branches and re-certify
# their actual command paths. Record hashes bind receipts, never enable policy.
CALIBRATED_IK_SEEDS = [[163.62039271007563, 64.01735255223417, -67.25050650734438, 93.2331539551102, -90.00000000000001, -106.37960728992437], [-72.40715810734315, -20.66480267505412, -103.89758096136477, 124.56238363641887, 72.40715810734312, 0.0], [-58.553344176794326, -22.475689666466394, -101.12528805253322, 123.60097771899962, 58.55334417679429, -1.0294949594003553e-14], [-58.553344176794326, -22.475689666466394, -101.12528805253322, 123.60097771899962, 58.55334417679429, 180.0], [-87.40476475829131, -22.47568966646641, -101.12528805253322, 123.60097771899962, 87.40476475829125, 180.0], [-64.66430037296594, -3.2481937678895747, -126.71804809984242, 129.96624186773198, 64.66430037296595, 180.0], [-75.41679324948196, -12.462263518678185, -56.77419042193441, -20.76354605938741, 90.0, 194.58320675051806], [-78.10373775148642, -37.83824919659381, -16.865010237740023, -35.296740565666134, 90.0, 191.89626224851355], [-88.23587605840977, -43.75520866199254, -5.060724146438354, -41.184067191569056, 90.0, 181.7641239415902], [-88.23587605840977, -43.75520866199254, -5.060724146438354, -41.184067191569056, 90.0, 1.7641239415902135], [-68.33462268250656, -43.75520866199333, -5.060724146436616, -41.184067191570016, 89.99999999999999, 21.665377317493437], [61.81374704354286, 48.51918849734889, 55.392423259627606, -103.91161175697648, 28.186252956457167, 180.0], [62.25330564679723, 54.06615976151417, 44.56648765802543, -98.6326474195396, 27.746694353202802, 180.0], [61.81374704354286, 48.51918849734889, 55.392423259627606, -103.91161175697648, 28.186252956457167, 90.0], [62.253305646797244, 54.06615976151415, 44.56648765802541, -98.63264741953954, 27.746694353202788, 89.99999999999999], [61.81374704354286, 48.51918849734889, 55.392423259627606, -103.91161175697648, 28.18625295645714, -90.00000000000001], [62.25330564679723, 54.0661597615141, 44.56648765802556, -98.63264741953965, 27.746694353202773, -90.00000000000004], [62.57433490659918, 47.78974891048301, 57.14855554302247, -103.76676871515006, 27.416346223420135, -60.70732349501101], [62.98154845233014, 53.155168153175346, 46.7150047327387, -98.68233310181975, 27.009218983764953, -60.72565665513798], [62.57582549469282, 48.080389017894106, 56.23528280269005, -104.31567182058413, 27.424174505307207, -180.0], [62.71034615480792, 51.83128832842894, 49.315963732196764, -99.89133677590429, 25.437207443150072, -301.4668568689523], [60.218467190004304, 39.42913510297621, 54.58098026787218, -92.8583848548389, 27.92853761288419, -301.35028218541504], [-13.591622773947876, 18.9460252211274, 48.02925373146127, 23.02472104741136, -90.0, -193.59162277394785]]
_continuous_profile_active = False


def _records_fingerprint(records):
    import hashlib
    canonical = [dict(type=r['type'], values=[0.0 if abs(float(v)) < 1e-12 else float(v)
                 for v in r['values']], singular=bool(r.get('singular', False)),
                 spin360=bool(r.get('spin360', False)), j6_delta=int(r.get('j6_delta', 0)))
                 for r in records]
    return hashlib.sha256(json.dumps(canonical, sort_keys=True,
        separators=(',', ':')).encode('utf-8')).hexdigest()


def _continuous_records(records):
    return len(records) > 1 and any(r.get('type') == 'TCP' for r in records)


def _assert_continuous_dispatch(records, initial, plan, direct_enabled):
    if not _continuous_records(records):
        return
    fingerprint = _records_fingerprint(records)
    previous = initial
    for number, step in enumerate(plan, 1):
        if step.get('waypoints'):
            certificate = step.get('direct_certificate') or {}
            if (step['method'] != 'MoveL' or not step.get('direct_movl_certified')
                    or certificate.get('records_sha256') != fingerprint
                    or certificate.get('start_joints') != list(previous)
                    or certificate.get('end_joints') != step['joints']
                    or certificate.get('send_joints') != step.get('direct_send_joints')):
                raise RuntimeError(f'P{number}缺少与当前数据及构型一致的连续直线认证，禁止退回逐点停走。')
            if not direct_enabled:
                raise RuntimeError('连续TCP轨迹需要单条MovL模式，禁止退回细分停走。')
        previous = step['joints']


def _controller_body_matches():
    expected = Fanuc_2_Pose([1.119989104069524, -245.1846134160959,
        1047.9330384567963, -89.7671431696512, -0.00006721956284782927,
        179.8638590144166])
    err = invH(expected) * robot.SolveFK([0.0] * 6)
    return norm(err.Pos()) < .001 and pose_angle(err) < math.radians(.001)


def _profile_ik_all(flange):
    native = robot.SolveIK_All(flange)
    if not _continuous_profile_active:
        return native
    key = ('profile_ik', _cache_key_pose(flange))
    if key in _plan_cache:
        return _plan_cache[key]
    raw = [list(q[:6]) for q in native]
    for seed in CALIBRATED_IK_SEEDS:
        q = robot.SolveIK(flange, seed).list()
        if len(q) >= 6:
            raw.append(q[:6])
    valid = []
    for q in raw:
        if len(q) != 6:
            continue
        q = [(float(v) + 180.0) % 360.0 - 180.0 for v in q]
        err = invH(flange) * robot.SolveFK(q)
        if norm(err.Pos()) > .001 or pose_angle(err) > math.radians(.001):
            continue
        if not any(max(abs(x-y) for x, y in zip(q, old)) < .001 for old in valid):
            valid.append(q)
    result = Mat(valid).tr() if valid else Mat(6, 0)
    _plan_cache[key] = result
    return result


def _direct_step_allowed(number, step):
    return number not in MOVL_DIRECT_BLOCK_POINTS or bool(step.get('direct_movl_certified'))


def _certify_continuous_direct(records, initial, plan, log):
    if not _continuous_profile_active:
        return
    if RDK.RunMode() != RUNMODE_SIMULATE or not _controller_body_matches():
        raise RuntimeError('本体或模式与连续TCP单条MovL验证条件不一致。')
    pose, link, frame, saved = robot.PoseTool(), robot.getLink(ITEM_TYPE_TOOL), robot.PoseFrame(), robot.Joints().list()[:6]
    lower, upper, _ = robot.JointLimits()
    try:
        for number, step in enumerate(plan, 1):
            if step['method'] != 'MoveL':
                continue
            if step['method'] != 'MoveL' or not step.get('waypoints'):
                raise ValueError(f'P{number}未形成连续直线，禁止以MoveJ代替本次工艺段。')
            start = initial if number == 1 else plan[number-2]['joints']
            relative = _trajectory_pose(step['joints']) * invH(_trajectory_pose(start))
            if norm(relative.Pos()) > MOVL_DIRECT_MAX_MM or pose_angle(relative) > math.radians(.5):
                raise ValueError(f'P{number}将退回{len(step["waypoints"])}段停走，换入口分支重试。')
            send_q, note = _movl_digit_safe_joints(step['joints'])
            if send_q is None:
                raise ValueError(f'P{number}发送位姿净化失败。')
            target = invH(frame) * robot.SolveFK(send_q)
            flange_tool = _named_tool(FLANGE_TOOL_NAME, eye(4))
            robot.setPoseTool(flange_tool)
            robot.setJoints(start)
            if robot.MoveL_Test(start, target, minstep_mm=.5) != 0:
                raise ValueError(f'P{number}净化后的法兰直线碰撞或不可达。')
            program = RDK.AddProgram('_轨迹16_单条MovL复核', robot)
            try:
                program.setVisible(False)
                program.setPoseTool(eye(4))
                program.setPoseFrame(frame)
                program.MoveJ(start)
                program.MoveL(send_q)
                robot.setJoints(start)
                message, matrix, status = program.InstructionListJoints(
                    mm_step=.5, deg_step=.2, collision_check=COLLISION_ON)
                samples = matrix.tr().rows
                if status < 0 or 'collision' in message.lower() or not samples:
                    raise ValueError(f'P{number}法兰整段复核失败：{message}')
                for row in samples:
                    q = row[:6]
                    if (int(row[6]) != 0 or not _real_limit_ok(q, lower.list(), upper.list())
                            or _real_interfere_combo(q)):
                        raise ValueError(f'P{number}法兰路径存在错误、限位或自干涉。')
                if max(abs(a-b) for a, b in zip(samples[-1][:6], send_q)) > .05:
                    raise ValueError(f'P{number}法兰直线落点分支与认证关节不一致。')
                err = invH(robot.SolveFK(send_q)) * robot.SolveFK(samples[-1][:6])
                if norm(err.Pos()) > .01 or pose_angle(err) > math.radians(.01):
                    raise ValueError(f'P{number}法兰路径终点不匹配。')
                step['direct_movl_certified'] = True
                step['direct_send_joints'] = list(send_q)
                step['direct_certificate'] = dict(records_sha256=_records_fingerprint(records),
                    start_joints=list(start), end_joints=list(step['joints']), send_joints=list(send_q),
                    samples=len(samples), flange_target=Pose_2_Fanuc(target), digit_note=note)
                log(f'P{number}：单条法兰MovL复核通过（0.5mm采样、碰撞/实机限位/落点分支）；本次免除细分。')
            finally:
                program.Delete()
                _restore_tool(pose, link)
    finally:
        _restore_tool(pose, link)
        robot.setPoseFrame(frame)
        robot.setJoints(saved)


def _ik_branch_candidates(target_pose, reference):
    """v14c：某个 TCP 位姿的全部限位内 IK 分支（含 J6 圈数取近表示），
    与 _nearest_ik_from_current 同款筛选规则。"""
    solutions = _profile_ik_all(_tcp_target_to_flange(target_pose))
    lower, upper, _ = robot.JointLimits()
    lower, upper = lower.list(), upper.list()
    candidates = []
    for solution in solutions:
        q = [((float(v) + 180.0) % 360.0) - 180.0 for v in solution[:6]]
        if len(q) != 6:
            continue
        for turns6 in (0, -1, 1):
            candidate = q[:]
            candidate[5] += 360.0 * turns6
            if _real_limit_ok(candidate, lower, upper):
                if not any(max(abs(a-b) for a, b in zip(candidate, old)) < 1e-6 for old in candidates):
                    candidates.append(candidate)
    for q in candidates[:]:
        nearest = [min((v + 360*k for k in range(math.ceil((lower[j]-v)/360),
                       math.floor((upper[j]-v)/360)+1)), key=lambda a: abs(a-reference[j]))
                   for j, v in enumerate(q)]
        # v14w22：取近表示必须复核实机限位（此前漏检 ⇒ J1=193.59 混入实发被 -40001 拒）
        if not _real_limit_ok(nearest, lower, upper):
            continue
        if not any(max(abs(a-b) for a, b in zip(nearest, old)) < 1e-6 for old in candidates):
            candidates.append(nearest)
    return candidates


def _nearest_ik_from_current_lookahead(current_q, target_pose, lookahead_ok):
    """v14i：同 _nearest_ik_from_current，但要求选出的解能满足前视条件 lookahead_ok(cand)->bool；
    没有满足者时退回最近解（死路由后续救援链/种子重试兜底）。"""
    candidates = _ik_branch_candidates(target_pose, current_q)
    if not candidates:
        raise ValueError('没有限位内的逆解。')
    ranked = sorted(candidates, key=lambda q: sum((q[j]-current_q[j])**2 for j in range(6)))
    for cand in ranked:
        if lookahead_ok(cand):
            return cand[:]
    return ranked[0][:]


def _nearest_ik_from_current(current_q, target_pose):
    """v14-P2P：从全部逆解中选离当前关节角最近的解（含 J6 圈数取近）。

    与 test.py 的肘高排序不同：以【关节空间离当前构型最近】为准，相邻点之间不会突变构型。
    没有限位内解时抛 ValueError。"""
    solutions = _profile_ik_all(_tcp_target_to_flange(target_pose))
    lower, upper, _ = robot.JointLimits()
    lower, upper = lower.list(), upper.list()
    candidates = []
    for solution in solutions:
        q = [((float(v) + 180.0) % 360.0) - 180.0 for v in solution[:6]]
        if len(q) != 6:
            continue
        for turns6 in (0, -1, 1):
            candidate = q[:]
            candidate[5] += 360.0 * turns6
            if _real_limit_ok(candidate, lower, upper):
                if not any(max(abs(a-b) for a, b in zip(candidate, old)) < 1e-6 for old in candidates):
                    candidates.append(candidate)
    # 同一姿态再补一圈数取近的表示，避免强制归零导致大绕行。
    for q in candidates[:]:
        nearest = [min((v + 360*k for k in range(math.ceil((lower[j]-v)/360),
                       math.floor((upper[j]-v)/360)+1)), key=lambda a: abs(a-current_q[j]))
                   for j, v in enumerate(q)]
        # v14w22：取近表示必须复核实机限位（此前漏检 ⇒ J1=193.59 混入实发被 -40001 拒）
        if not _real_limit_ok(nearest, lower, upper):
            continue
        if not any(max(abs(a-b) for a, b in zip(nearest, old)) < 1e-6 for old in candidates):
            candidates.append(nearest)
    if not candidates:
        raise ValueError('没有限位内的逆解。')
    return min(candidates, key=lambda q: sum((q[j]-current_q[j])**2 for j in range(6)))[:]


def _checked_j6_rewinds(q, lower, upper, max_deviation):
    """返回可实际执行的整圈回绕列表（带缓存）；TCP空间偏离和碰撞都必须通过检查。"""
    key = ('rewinds', _cache_key_joints(q), tuple(round(float(v), 6) for v in lower[:6]),
           tuple(round(float(v), 6) for v in upper[:6]), round(float(max_deviation), 6))
    if key in _plan_cache:
        return [r[:] for r in _plan_cache[key]]
    results = []
    tcp = pose_to_fanuc_values(_trajectory_pose(q))
    for delta in (-360.0, 360.0):
        end = q[:]
        end[5] += delta
        if not lower[5] <= end[5] <= upper[5]:
            continue
        if not _check_movej_tcp_trajectory(q, end, tcp, tcp, lambda msg: None,
                                          samples=360, max_deviation_mm=max_deviation):
            continue
        if _movej_test_cached(q, end, 1) == 0:
            results.append(end)
    _plan_cache[key] = results
    return [r[:] for r in results]


def _plan_continuous_trajectory(records, max_deviation, log):
    """v14c：首点全分支种子枚举 + 整段重试。

    贪心最近解在换向步（如轨迹7 P6 的原地转 90°→180°）会把 wrist 构型选到贴圆柱，
    后续任何分支都碰；TCP仿真宏靠首点种子枚举+整段重试避开这类死路。v14c 移植该机制：
    种子按肘高排序优先，贪心只负责段内选解；某段死路（含 MoveL 兑底都失败）
    则整段换种子重试，全部种子失败才报错。"""
    global _preferred_seed, _continuous_profile_active
    _continuous_profile_active = False
    if _continuous_records(records):
        if not _controller_body_matches():
            raise RuntimeError('连续TCP轨迹策略要求控制器对齐本体；当前本体参数不符。')
        if not _same_tool_pose(robot.PoseTool(), Fanuc_2_Pose(list(CANONICAL_TOOL))):
            raise RuntimeError('连续TCP轨迹策略要求130mm TCP。')
        if norm(robot.PoseFrame().Pos()) > .01 or pose_angle(robot.PoseFrame()) > math.radians(.01):
            raise RuntimeError('连续TCP轨迹策略要求机器人基座参考系。')
        _continuous_profile_active = True
        log('v15.21：启用校准本体分支搜索及防停走检查；不依赖旧坐标指纹，全部直线按当前数据重新认证。')
    _enable_obstacle_checks()
    if not math.isfinite(max_deviation) or max_deviation < 0:
        raise ValueError('MoveJ允许偏离必须是非负有限数。')
    for i, rec in enumerate(records):
        vals = rec['values']
        if rec['type'] not in ('TCP', 'JOINT') or len(vals) != 6 or not all(math.isfinite(v) for v in vals):
            raise ValueError(f'P{i+1}：点类型或六维数值无效。')
        if rec.get('singular', False):
            # v14a：恢复 v13 同款奇异点规则校验（P2P 规划层支持奇异点步）
            if rec['type'] != 'TCP' or i == 0 or records[i-1]['type'] != 'TCP' or records[i-1].get('singular', False):
                raise ValueError(f'P{i+1}：特异点必须紧跟普通TCP点。')
            if rec.get('spin360', False):
                if rec.get('j6_delta', 360) not in (-360, 360):
                    raise ValueError(f'P{i+1}：J6自转方向必须为+360或-360。')
                if max(abs(a - b) for a, b in zip(rec['values'], records[i-1]['values'])) > 1e-3:
                    raise ValueError(f'P{i+1}：J6自转360°特异点的六维数值必须与前一个TCP点完全相同。')
            elif rec.get('j6_delta', 180) not in (-180, 180):
                raise ValueError(f'P{i+1}：J6方向必须为+180或-180。')
    saved = robot.Joints().list()[:6]
    lower, upper, _ = robot.JointLimits()
    lower, upper = lower.list(), upper.list()
    # 先检查点本身可达，避免后面的不可达点触发整段分支重复搜索。
    unreachable = []
    for i, rec in enumerate(records, 1):
        if rec['type'] == 'TCP' and not rec.get('singular', False):
            target = fanuc_values_to_pose(*rec['values'])
            if _profile_ik_all(_tcp_target_to_flange(target)).size(1) == 0:
                unreachable.append(f'P{i}：没有逆解；' + _flange_target_description(target))
    if unreachable:
        raise ValueError('目标点不可达，尚未搜索连接路径：' + '；'.join(unreachable))
    if _movej_test_cached(saved, saved, 1) != 0:
        raise ValueError('起始姿态已碰撞，不能自动规划脱离：' + _collision_details())
    try:
        RDK.Render(False)
        # v14c：首点全分支种子枚举（肘高优先），某种子整段死路时换构型重试。
        first_tcp = next((r for r in records if r['type'] == 'TCP' and not r.get('singular', False)), None)
        if first_tcp is not None:
            seeds = _ik_branch_candidates(fanuc_values_to_pose(*first_tcp['values']), saved)
            seeds.sort(key=lambda s: _obstacle_posture_key(s, saved))
            if _continuous_profile_active:
                # Recover the previously successful entry branch on this calibrated body.
                # These are IK seeds, never executable joint targets.
                entry = robot.SolveIK(_tcp_target_to_flange(
                    fanuc_values_to_pose(*first_tcp['values'])), CALIBRATED_IK_SEEDS[0]).list()
                if len(entry) == 6:
                    seeds.sort(key=lambda s: sum((a-b)**2 for a,b in zip(s, entry)))
                log('v15.21：优先历史成功入口分支；任何细分停走退化均重新选解或停止预检。')
        else:
            seeds = [None]
        seed_context = repr((records, saved, robot.PoseFrame().rows, robot.PoseTool().rows, max_deviation))
        if _preferred_seed is not None and _preferred_seed[0] == seed_context:
            preferred = _preferred_seed[1]
            seeds.sort(key=lambda s: 0 if s == preferred else 1)
            log('优先尝试上次通过的首点构型；本次所有碰撞与整段检查仍重新执行。')
        last_seed_error = None
        for seed_rank, seed in enumerate(_lazy_valid_seeds(seeds, saved), 1):
            if len(seeds) > 1:
                log(f'—— 尝试首点分支种子 {seed_rank}/{len(seeds)}：' +
                    ('%s' % [round(v, 1) for v in seed] if seed else '无种子(关节轨迹)'))
            q = saved[:]
            plan = []
            try:
                seed_used = seed is None
                for i, rec in enumerate(records, 1):
                    rewinds = []
                    delta = None
                    method, fallback, waypoints = 'MoveJ', False, []
                    lookahead_ok = None  # v14j：循环顶初始化（首个TCP点走种子路径时前视绑定也可安全引用）
                    if rec['type'] == 'JOINT':
                        end = [float(v) for v in rec['values'][:6]]
                        note = '录入关节直达'
                    elif rec.get('singular', False):
                        # v14a：奇异点步——只转 J6（±180 换向 / ±360 自转）。
                        # ±180：从当前解纯转 J6，由下方 FK 校验把关；超限时先试反方向（终点位姿不变）再试整圈回绕。
                        target = fanuc_values_to_pose(*rec['values'])
                        delta = rec.get('j6_delta', 180)

                        def _fk_matches(candidate):
                            error_pose = invH(target) * _trajectory_pose(candidate)
                            return norm(error_pose.Pos()) <= 1e-3 and pose_angle(error_pose) <= math.radians(.01)

